(* IEC 61131-3 sources: daoli-st-library/DL_Motion, 205 files *)

(* ---- FB_DL_AxisBacklashIdent.st ---- *)
(*==============================================================================
 * 组件名称 (Component)  : FB_DL_AxisBacklashIdent
 * 所属子库 (Sublibrary) : DL_Motion
 * 当前版本 (Version)    : 1.0.0
 * 兼容性   (Platform)   : CODESYS 3.5+ / TwinCAT 3 / 汇川 InoProShop / 施耐德 Machine Expert
 *                         仅依赖 Standard.library（R_TRIG），零厂商私有库
 * 功能描述 (Function)   : 反向间隙在线辨识（只辨识、不注入）。
 *                         原理：换向瞬间传动链要"先吃掉间隙"才带动负载，故换向后的**指令位移**与
 *                         **实际位移**之差即间隙的一次观测值。本件在每个换向沿开启一个位移窗，
 *                         窗内位移超过 fWinMoveMm 即结算一个残差样本：
 *                           残差 = | (Δ指令位移) − (Δ实际位移) | [mm]
 *                         样本进定长缓冲（8 个），样本数达 nMinSamples 后取**中值**作为间隙估计
 *                         （中值对个别打滑/编码器毛刺样本免疫，均值则不）。
 *                         三条固化纪律：
 *                           ① **激励不足拒辨识**：样本数不足或换向时速度幅值低于 fVelMin 时，
 *                              估计值不宣称（bValid=FALSE）并置 bInsufficientExc——低速换向的残差
 *                              被摩擦完全淹没，硬算出来的"间隙"只是摩擦的另一种写法；
 *                           ② **中值估计**：样本排序后取中位（8 个样本插入排序，循环上界恒定）；
 *                           ③ **估计值钳位**：结果钳 [0, fBacklashMax]，超上限按上限报告并置 bClamped
 *                              （不可信的巨值不许直接进入补偿环节）。
 *                         验收向量：
 *                           ① 五次换向残差 {0.02, 0.03, 0.03, 0.04, 0.10} → 中值 0.03 mm（0.10 为野值）
 *                           ② 仅 2 个样本（nMinSamples=5）→ bValid=FALSE + bInsufficientExc
 *                           ③ 换向时速度 0.5 mm/s（fVelMin=2.0）→ 该次不采样本
 *                           ④ 残差 5.0 mm（上限 2.0）→ 估计钳 2.0 mm + bClamped
 * 接口     (Interface)  : 入 bEnable 使能、fCmdPos 指令位置、fActPos 实际位置、fVelCmd 指令速度、
 *                         fVelMin 换向速度下限（激励门槛）、fWinMoveMm 位移窗宽、fBacklashMax 估计上限、
 *                         nMinSamples 最少样本数（≥1）、bClear 清样本沿、bReset 复位沿；
 *                         出 fBacklashMm 间隙估计（中值）、bValid 估计有效、bClamped 估计被钳位、
 *                         iSampleCnt 已收样本数、bInsufficientExc 激励不足、bReversed 换向脉冲（单拍）、
 *                         eState 相、eCause 成因、bError 故障标志。
 * 边界     (Boundary)   : ① **属主边界（写死）：本件只做"间隙辨识"，不注入补偿、不改位置环输出**——
 *                         补偿注入属上层（`FB_DL_AxisCoggingFf` 族与本件并列不互引）；
 *                         ② **状态枚举禁定义**：本件不引用任何轴状态枚举（R277），只消费位置/速度引脚；
 *                         ③ **组态闸**：fVelMin > 0、fWinMoveMm > 0、fBacklashMax > 0、nMinSamples ≥ 1
 *                         且 ≤ 8，违反即锁存 eCfgIllegal；
 *                         ④ **非有限闸**：任一位置/速度样本非有限 → 该拍不采样（不锁存）；
 *                         ⑤ **样本缓冲边界**：8 样本字面量上界（R104），写入前判满；
 *                         ⑥ **锁存解除式**：eFault 仅由 bReset 上升沿解除（R228B），bReset 恒可达；
 *                         ⑦ 零全局耦合、零物理地址。
 * 分工声明 (Scope)      : 本件只管"换向残差统计与中值估计"。不接管：摩擦前馈
 *                         （属 FB_DL_AxisFrictionFf）、齿槽前馈（属 FB_DL_AxisCoggingFf）、
 *                         双反馈切换（属 AxisFeedbackFailoverSeq 族）。
 * 来源标签 (Source Tag) : 自研线（传动精度族开族）
 * 码表     (Codes)      : 本件不占用任何全局数字码位（零码位范式 R297）；诊断由 BOOL + ENUM 出口承担。
 * 红线自检 (Redline)    : R1 ✓ 零 GVL/VAR_EXTERNAL ｜ R2 ✓ 零 %I/%Q/%M ｜ R3 ✓ 纯 IEC 61131-3
 *                         R4 ✓ 组态闸 + 非有限闸 + 缓冲边界 + 估计钳位 ｜ R5 ✓ 声明逐行同行双语注释
 *                         R6 ✓ ENUM+CASE 含 ELSE 兜底 ｜ R7 ✓ 三 R_TRIG 段 0 无条件刷新（本件无 TON）
 * 修订历史 (Revision)   : 2026-11-19  v1.0.0  R47 首版（批次 4 · 序号 19）
 *==============================================================================*)

TYPE E_DL_AbiState :
(
    eIdle  := 0,    // 待机相（未使能或已清零） / Idle, disabled or cleared
    eWatch := 10,   // 观测相（等换向沿并结算样本） / Watching, awaiting reversal and sample settlement
    eFault := 90    // 故障相（组态非法，等复位） / Fault, awaiting reset
);
END_TYPE

TYPE E_DL_AbiCause :
(
    eNone           := 0,   // 无异常 / No anomaly
    eCfgIllegal     := 1,   // 组态非法（门槛/窗口/上限/样本数越域） / Illegal configuration
    eInsufficientExc:= 2,   // 激励不足（样本数不够或换向速度过低） / Insufficient excitation
    eClamped        := 3,   // 估计值被钳位（野值） / Estimate clamped
    eSampleBad      := 4,   // 位置/速度样本非有限（当拍不采） / Non-finite sample, skipped
    ePhaseBad       := 5    // 非法相位兜底 / Illegal phase fallback
);
END_TYPE

FUNCTION_BLOCK FB_DL_AxisBacklashIdent
VAR_INPUT
    bEnable      : BOOL := FALSE;      // 使能（FALSE 冻结观测，不宣称） [-] / Enable
    fCmdPos      : LREAL := 0.0;       // 指令位置 [mm] / Command position [mm]
    fActPos      : LREAL := 0.0;       // 实际位置 [mm] / Actual position [mm]
    fVelCmd      : LREAL := 0.0;       // 指令速度（用于换向判定） [mm/s] / Command velocity [mm/s]
    fVelMin      : LREAL := 2.0;       // 换向速度下限（激励门槛），域 > 0 [mm/s] / Reversal speed limit, > 0
    fWinMoveMm   : LREAL := 1.0;       // 位移窗宽，域 > 0 [mm] / Displacement window, > 0
    fBacklashMax : LREAL := 2.0;       // 估计上限，域 > 0 [mm] / Estimate ceiling, > 0
    nMinSamples  : INT := 5;           // 最少样本数，域 1..8 [个] / Minimum sample count, 1..8
    bClear       : BOOL := FALSE;      // 清样本沿（重新辨识） [-] / Clear-samples edge
    bReset       : BOOL := FALSE;      // 故障复位沿 [-] / Fault reset edge
END_VAR
VAR_OUTPUT
    fBacklashMm   : LREAL := 0.0;                        // 间隙估计（中值，已钳位） [mm] / Backlash estimate, clamped
    bValid        : BOOL := FALSE;                       // 估计有效（样本够且激励足） [-] / Estimate valid
    bClamped      : BOOL := FALSE;                       // 估计被钳位 [-] / Estimate clamped
    iSampleCnt    : INT := 0;                            // 已收样本数 [个] / Collected sample count
    bInsufficientExc : BOOL := FALSE;                    // 激励不足 [-] / Insufficient excitation
    bReversed     : BOOL := FALSE;                       // 换向脉冲（单拍） [-] / Reversal pulse, single scan
    eState        : E_DL_AbiState := E_DL_AbiState.eIdle;    // 相出口 [-] / Phase outlet
    eCause        : E_DL_AbiCause := E_DL_AbiCause.eNone;    // 成因出口（R190 归因唯一） [-] / Cause outlet
    bError        : BOOL := FALSE;                       // 故障标志（仅组态级） [-] / Error flag, configuration only
END_VAR
VAR
    _eState   : E_DL_AbiState := E_DL_AbiState.eIdle;    // 内部相（CASE 唯一写入目标） / Internal phase
    _eCause   : E_DL_AbiCause := E_DL_AbiCause.eNone;    // 成因锁存量 / Latched cause
    _bFault   : BOOL := FALSE;                           // 故障锁存位 / Latched fault bit
    _iCnt     : INT := 0;                                // 样本计数 / Sample count
    _bDirPos  : BOOL := FALSE;                           // 上拍方向为正标志 / Previous direction positive flag
    _bDirNow  : BOOL := FALSE;                           // 当拍方向标志 / Present direction flag
    _bWinOpen : BOOL := FALSE;                           // 位移窗开启标志 / Displacement window open
    _fCmdSnap : LREAL := 0.0;                            // 换向瞬间指令位置快照 [mm] / Command snapshot at reversal
    _fActSnap : LREAL := 0.0;                            // 换向瞬间实际位置快照 [mm] / Actual snapshot at reversal
    _fResid   : LREAL := 0.0;                            // 残差工作值 [mm] / Residual working value
    _fEst     : LREAL := 0.0;                            // 中值估计工作值 [mm] / Median working value
    _fTmp     : LREAL := 0.0;                            // 排序交换临时量 [mm] / Sort swap temporary
    _bRev     : BOOL := FALSE;                           // 换向脉冲内部位（单拍） / Internal reversal pulse
    _bClamped : BOOL := FALSE;                           // 钳位标志内部位 / Internal clamp flag
    _bSampleOk: BOOL := FALSE;                           // 样本有限性结论 / Sample finiteness result
    _bCfgBad  : BOOL := FALSE;                           // 组态非法当拍量 / Illegal configuration this scan
    _i        : INT := 0;                                // 样本循环下标 / Sample loop index
    _j        : INT := 0;                                // 排序内层下标 / Inner sort index
    rtClear   : R_TRIG;                                  // 清样本沿实例，段 0 无条件调用 / Clear edge instance
    rtReset   : R_TRIG;                                  // 复位沿实例，段 0 无条件调用 / Reset edge instance
    afSmp     : ARRAY[1..8] OF LREAL;                    // 残差样本缓冲（字面量上界，R104） [mm] / Residual sample buffer
    afSort    : ARRAY[1..8] OF LREAL;                    // 排序副本 [mm] / Sorting copy
END_VAR
VAR CONSTANT
    DL_ABI_NMAX : INT := 8;            // 样本缓冲深度（与数组字面量上界同源） [个] / Sample buffer depth
    DL_ABI_EPS  : LREAL := 1.0E-12;    // 浮点判等容差 [mm] / Equality tolerance
END_VAR

(* —— 段 0：组态闸 + 三沿无条件周期刷新（R228A；本件无 TON） —— *)
_bCfgBad := (fVelMin <= 0.0) OR (fWinMoveMm <= 0.0) OR (fBacklashMax <= 0.0)      // 三正域闸 / Three positive-domain gates
         OR (nMinSamples < 1) OR (nMinSamples > DL_ABI_NMAX);                     // 样本数域闸 / Sample count domain
rtClear(CLK := bClear);                                                            // 清样本沿 / Clear edge
rtReset(CLK := bReset);                                                            // 复位沿 / Reset edge

(* —— 段 1：单拍/输出量预置（锁存量 _eCause/_bFault/_iCnt/_bWinOpen/_bDirPos 不入清单，R107） —— *)
bValid   := FALSE;                                                                 // 有效位预置 / Validity preset
_bRev    := FALSE;                                                                 // 换向脉冲预清 / Reversal pulse preset
_bClamped:= FALSE;                                                                 // 钳位标志预清 / Clamp flag preset
bInsufficientExc := FALSE;                                                         // 激励不足预清 / Insufficient-excitation preset
bError   := FALSE;                                                                 // 故障标志预清（R45 配对） / Error preset
_fEst    := 0.0;                                                                   // 估计工作值预置 / Estimate preset

(* —— 段 2：组态闸（非法即锁存） —— *)
IF _bCfgBad THEN
    _eCause := E_DL_AbiCause.eCfgIllegal;                                          // 归因：组态非法 / Cause: illegal configuration
    _bFault := TRUE;                                                               // 锁存 / Latch
    _eState := E_DL_AbiState.eFault;                                               // 入故障相 / Enter fault phase
END_IF

(* —— 段 3：迁出链与清样本链（两条显式写出） —— *)
IF rtReset.Q THEN
    _bFault   := FALSE;                                                            // 清故障锁存 / Clear fault latch
    _eCause   := E_DL_AbiCause.eNone;                                              // 清成因 / Clear cause
    _iCnt     := 0;                                                                // 样本清零 / Samples cleared
    _bWinOpen := FALSE;                                                            // 关窗 / Window closed
    _eState   := E_DL_AbiState.eIdle;                                              // 回待机相 / Back to idle
END_IF
IF rtClear.Q THEN
    _iCnt     := 0;                                                                // 样本清零（重新辨识） / Samples cleared for re-identification
    _bWinOpen := FALSE;                                                            // 关窗 / Window closed
END_IF

(* —— 段 4：相迁移（使能驱动；故障相由段 3 迁出） —— *)
CASE _eState OF

E_DL_AbiState.eIdle:
    IF bEnable AND (NOT _bCfgBad) THEN
        _eState := E_DL_AbiState.eWatch;                                           // 使能进观测相 / Enter watching
    END_IF

E_DL_AbiState.eWatch:
    IF NOT bEnable THEN
        _eState := E_DL_AbiState.eIdle;                                            // 失能回待机相（不借故障相过桥，R211） / Back to idle
    END_IF

E_DL_AbiState.eFault:
    ;                                                                              // 故障相：由段 3 复位沿迁出 / Exit via the reset edge

ELSE
    _eCause := E_DL_AbiCause.ePhaseBad;                                            // 归因：非法相位 / Cause: illegal phase
    _bFault := TRUE;                                                               // 锁存 / Latch
    _eState := E_DL_AbiState.eFault;                                               // 强拉故障相 / Force fault phase

END_CASE

(* —— 段 5：换向检测与窗结算（样本采集唯一入口） —— *)
IF _eState = E_DL_AbiState.eWatch THEN
    _bSampleOk := NOT ((fCmdPos <> fCmdPos) OR ((fCmdPos - fCmdPos) <> (fCmdPos - fCmdPos)))
              AND NOT ((fActPos <> fActPos) OR ((fActPos - fActPos) <> (fActPos - fActPos)))
              AND NOT ((fVelCmd <> fVelCmd) OR ((fVelCmd - fVelCmd) <> (fVelCmd - fVelCmd)));

    IF _bSampleOk THEN
        (* 换向判定：速度符号翻转且幅值过激励门槛；方向保持量只在激励充分时更新 *)
        _bDirNow := (fVelCmd > 0.0);                                               // 本拍方向 / Present direction
        IF (ABS(fVelCmd) > fVelMin) THEN
            IF (_bDirNow <> _bDirPos) AND (NOT _bWinOpen) THEN
                _bRev     := TRUE;                                                 // 换向脉冲（内部位） / Internal reversal pulse
                _bWinOpen := TRUE;                                                 // 开位移窗 / Open the displacement window
                _fCmdSnap := fCmdPos;                                              // 记录指令基准 / Command snapshot
                _fActSnap := fActPos;                                              // 记录实际基准 / Actual snapshot
            END_IF
            _bDirPos := _bDirNow;                                                  // 方向保持量更新 / Refresh the direction
        END_IF

        (* 窗结算：指令位移超过窗宽即结算一个残差样本 *)
        IF _bWinOpen AND (ABS(fCmdPos - _fCmdSnap) > fWinMoveMm) THEN
            _fResid := ABS((fCmdPos - _fCmdSnap) - (fActPos - _fActSnap));         // 残差 = |Δ指令 − Δ实际| / Residual
            IF _fResid <> _fResid THEN
                _fResid := 0.0;                                                    // 残差非有限：拒收（不采样本） / Non-finite residual rejected
                _eCause := E_DL_AbiCause.eSampleBad;                               // 归因：样本非有限 / Cause: sample non-finite
            ELSIF _iCnt < DL_ABI_NMAX THEN
                _iCnt := _iCnt + 1;                                                // 样本计数 +1 / Sample count increment
                afSmp[_iCnt] := _fResid;                                           // 落样本（下标已判满） / Store the sample
            END_IF
            _bWinOpen := FALSE;                                                    // 关窗，等下次换向 / Close the window
        END_IF
    ELSE
        _eCause := E_DL_AbiCause.eSampleBad;                                       // 归因：样本非有限（当拍不采） / Cause: non-finite sample
    END_IF

    (* —— 段 6：中值估计（只对已收样本排序；插入排序，循环上界为样本数 ≤ 8） —— *)
    IF _iCnt >= nMinSamples THEN
        FOR _i := 1 TO _iCnt DO
            afSort[_i] := afSmp[_i];                                               // 复制已收样本 / Copy the collected samples
        END_FOR
        FOR _i := 2 TO _iCnt DO
            _j := _i;                                                              // 插入排序内层起点 / Insertion start
            WHILE (_j > 1) AND (afSort[_j - 1] > afSort[_j]) DO
                _fTmp := afSort[_j - 1];                                           // 交换 / Swap
                afSort[_j - 1] := afSort[_j];
                afSort[_j] := _fTmp;
                _j := _j - 1;                                                      // 内层推进（收敛，R74） / Inner step, converges
            END_WHILE
        END_FOR
        _fEst := afSort[(_iCnt / 2) + 1];                                          // 取中位（1 基，样本数 1..8） / Median, 1-based
        IF _fEst > fBacklashMax THEN
            _fEst := fBacklashMax;                                                 // 上限钳位（野值不许进入补偿） / Clamp to the ceiling
            _bClamped := TRUE;                                                     // 钳位标志 / Clamp flag
            _eCause := E_DL_AbiCause.eClamped;                                     // 归因：估计被钳位 / Cause: estimate clamped
        ELSIF _fEst < 0.0 THEN
            _fEst := 0.0;                                                          // 下限钳位（间隙非负） / Clamp to zero
            _bClamped := TRUE;                                                     // 钳位标志 / Clamp flag
            _eCause := E_DL_AbiCause.eClamped;                                     // 归因：估计被钳位 / Cause: estimate clamped
        END_IF
        bValid := TRUE;                                                            // 估计有效 / Estimate valid
    ELSE
        bInsufficientExc := TRUE;                                                  // 激励不足：不宣称 / Insufficient excitation
        _eCause := E_DL_AbiCause.eInsufficientExc;                                 // 归因：激励不足 / Cause: insufficient excitation
    END_IF
END_IF

(* —— 段 7：出口单点映射（名实双出口，R191） —— *)
fBacklashMm := _fEst;                                                              // 间隙估计出口 / Backlash estimate outlet
bClamped    := _bClamped;                                                          // 钳位标志出口 / Clamp flag outlet
iSampleCnt  := _iCnt;                                                              // 样本数出口 / Sample count outlet
bReversed   := _bRev;                                                              // 换向脉冲出口 / Reversal pulse outlet
eState      := _eState;                                                            // 相出口 / Phase outlet
eCause      := _eCause;                                                            // 成因出口 / Cause outlet
bError      := _bFault;                                                            // 故障标志 / Error flag

END_FUNCTION_BLOCK

(* ---- FB_DL_AxisFeedbackFailoverSeq.st ---- *)
(*==============================================================================
 * 组件名称 (Component)  : FB_DL_AxisFeedbackFailoverSeq
 * 所属子库 (Sublibrary) : DL_Motion
 * 当前版本 (Version)    : 1.0.1
 * 兼容性   (Platform)   : CODESYS 3.5+ / TwinCAT 3 / 汇川 InoProShop / 施耐德 Machine Expert
 *                         仅依赖 Standard.library（TON / R_TRIG / ABS），零厂商私有库
 * 功能描述 (Function)   : 主反馈（负载侧光栅尺/全闭环编码器）失效 → 电机侧反馈降级切换序。
 *                         四段序，每段语义显式，绝无"静默降级"：
 *                           ① ePrimary 主用相：bUsePrimary=TRUE，主反馈在岗；
 *                           ② eConfirm 失主确认相：主反馈有效位为假且持续 tLossConfirm；
 *                           ③ eSwitching 切换过渡相：**两侧均不宣称可用**（bUsePrimary 与
 *                              bUseMotorSide 同为假），先撤主用再等 tSwitchDwell，让轴级看到
 *                             一个明确的"无有效反馈"过渡拍，禁止无缝瞬切造成位置基准跳变；
 *                           ④ eDegraded 降级保持相：bUseMotorSide=TRUE 且 bFailoverActive 锁存置真，
 *                             告警持续可见直到人工复位（不因主反馈恢复而自动消失——那会让
 *                             维护人员永远看不到发生过降级）。
 *                         另设 eBlocked：主反馈已失效但 bSwitchPermit 为假（轴在运动中、
 *                         未到安全位）→ 置 bSwitchForbidden 告警，两侧反馈出口同为假，
 *                         交由轴级停机；**不做"先切了再说"**。
 * 接口     (Interface)  : 输入 bPrimaryValid 主反馈有效位、bSwitchPermit 允许切换（安全前置）、
 *                         tLossConfirm 失主确认时间、tSwitchDwell 切换过渡驻留时间、bReset 复位；
 *                         输出 bUsePrimary 用主反馈、bUseMotorSide 用电机侧、bFailoverActive
 *                         降级告警锁存、bSwitchForbidden 切换被禁止告警、eState / eCause / bError。
 * 边界     (Boundary)   : ① **属主边界（写死）：本件是"切换序"的唯一属主**——它决定何时撤主用、
 *                         何时上电机侧、过渡驻留多久。**判"负载侧是否可信"不是本件的职责**，
 *                         那属于 `FB_DL_AxisLoadEncoderLossMonitor`；本件只吃它的结论位
 *                         bPrimaryValid，不得内嵌断线/冻结判据（否则两件归因冲突、故障台账双记）。
 *                         ② 本件**不使能/不停止轴、不发运动指令**，只出反馈选择与告警位，
 *                         降级后的速度/位置环怎么跑由轴级 POU 决定。
 *                         ③ 组态闸：tLossConfirm <= T#0S → 故障锁存（防零时切换）。tSwitchDwell 的
 *                            "域 >= T#0S" 由类型本身保证（TIME 无符号），v1.0.1 已删除该恒假判据。
 *                         ④ 两枚 TON + 一枚 R_TRIG 段 0 无条件周期刷新，PT 语义成对写死；
 *                         切换过渡用 tonDwell（IN = 当拍位于 eSwitching），出相即 IN 落假自动复位，
 *                         无跨相累积（R228A）。
 *                         ⑤ 故障相与降级相均可迁出（R228B）：bReset 上升沿 → ePrimary。
 *                         ⑥ 零全局耦合（无 GVL / 无 VAR_EXTERNAL / 无物理地址）。
 * 分工声明 (Scope)      : 与 `FB_DL_AxisLoadEncoderLossMonitor`（只判负载侧可信度）、
 *                         `FB_DL_AxisDualFeedbackGuard`（双侧交叉校核）三件成组：监控件出结论，
 *                         本件按结论执行切换，校核件做一致性体检。三件互不内嵌对方判据。
 * 来源标签 (Source Tag) : P1 双反馈族 / T2-4 ◐
 * 解除式   (Release)    : bReset 上升沿（人工确认）→ 回 ePrimary 并清 bFailoverActive。
 *                         自证可满足：复位是外部操作员动作，不受任何锁存量门控；不设"主反馈自动
 *                         恢复即回切"的隐式路径——那会在反馈抖动时来回切换，且会抹掉降级告警痕迹。
 * 码表     (Codes)      : 本件不占用任何全局数字码位。出口为 BOOL（bUsePrimary / bUseMotorSide /
 *                         bFailoverActive / bSwitchForbidden / bError）+ ENUM（eState / eCause）；
 *                         数字码位待主控收口阶段统一派号（R46 码位规则）。
 * 红线自检 (Redline)    : R1 ✓ 零 GVL/VAR_EXTERNAL ｜ R2 ✓ 零 %I/%Q/%M ｜ R3 ✓ 纯 IEC 61131-3
 *                         R4 ✓ 时间域几何闸 + 无浮点比较 ｜ R5 ✓ 声明逐行同行双语注释
 *                         R6 ✓ ENUM+CASE 含 ELSE ｜ R7 ✓ TON/R_TRIG 段 0 无条件刷新
 * 返修记录 (Repair)     : v1.0.1（R47 P0 返修）① bError 出口增 `(_eState = eFault)` 项——原先只有禁止相
 *                         置位，故障相虽锁存却不报错，轴级不会停机；② 删除 `tSwitchDwell < T#0S` 恒假死检查
 *                         （TIME 为无符号时长量，与 0 的"小于"结构性不可达，属死判据）。
 * 修订历史 (Revision)   : 2026-11-19  v1.0.0  R46 首版（批次 2 · 序号 6）
 *==============================================================================*)

TYPE E_DL_FfsState :
(
    ePrimary   := 0,    // 主反馈在岗相 / Primary feedback in service
    eConfirm   := 10,   // 失主确认相（等 tLossConfirm） / Primary-loss confirmation
    eSwitching := 20,   // 切换过渡相（两侧均不宣称可用） / Switching transition, neither side claimed
    eDegraded  := 30,   // 降级保持相（电机侧在岗，告警锁存） / Degraded hold, alarm latched
    eBlocked   := 40,   // 切换被禁止相（安全前置未满足） / Switch forbidden phase
    eFault     := 90    // 组态故障相 / Configuration fault phase
);
END_TYPE

TYPE E_DL_FfsCause :
(
    eNone           := 0,   // 无故障成因 / No cause
    eCfgIllegal     := 1,   // 组态非法（确认时间非正/驻留为负） / Illegal configuration
    ePrimaryLost    := 2,   // 主反馈失效并已确认，完成降级 / Primary lost and confirmed, degraded
    eSwitchForbidden:= 3,   // 主反馈失效但切换前置不满足 / Primary lost but switching not permitted
    ePhaseBad       := 4    // 非法相位兜底 / Illegal phase fallback
);
END_TYPE

FUNCTION_BLOCK FB_DL_AxisFeedbackFailoverSeq
VAR_INPUT
    bPrimaryValid  : BOOL := TRUE;          // 主反馈（负载侧）有效位，来自监控件 [-] / Primary feedback validity, from the monitor unit
    bSwitchPermit  : BOOL := FALSE;         // 允许切换的安全前置（轴静止/在安全位） [-] / Safety precondition permitting the switch
    tLossConfirm   : TIME := T#100MS;       // 失主确认时间，域 > T#0S [ms] / Primary-loss confirm time, domain > T#0S
    tSwitchDwell   : TIME := T#20MS;        // 切换过渡驻留时间，域 >= T#0S [ms] / Switching dwell, domain >= T#0S
    bReset         : BOOL := FALSE;         // 人工复位，上升沿回主用相并清降级告警 [-] / Manual reset, rising edge returns to primary
END_VAR
VAR_OUTPUT
    bUsePrimary     : BOOL;     // 采用主反馈（负载侧） [-] / Use primary feedback
    bUseMotorSide   : BOOL;     // 采用电机侧反馈（降级后） [-] / Use motor-side feedback
    bFailoverActive : BOOL;     // 降级告警，锁存保持到复位（显式，不静默） [-] / Failover alarm, latched until reset
    bSwitchForbidden: BOOL;     // 切换被禁止告警（当拍量） [-] / Switch-forbidden alarm, per scan
    eState          : E_DL_FfsState;    // 状态出口 [-] / State outlet
    eCause          : E_DL_FfsCause;    // 成因出口（R190 归因唯一） [-] / Cause outlet
    bError          : BOOL;             // 故障标志（组态故障或切换被禁止） [-] / Error flag
END_VAR
VAR
    _eState    : E_DL_FfsState := E_DL_FfsState.ePrimary;    // 内部相位（CASE 唯一写入目标） / Internal phase
    _eCause    : E_DL_FfsCause := E_DL_FfsCause.eNone;       // 成因出口暂存（锁存语义由相位承载） / Cause staging
    tonLoss    : TON;           // 失主确认计时，段 0 无条件调用 / Primary-loss confirm timer
    tonDwell   : TON;           // 切换过渡驻留计时，段 0 无条件调用 / Switching dwell timer
    rtReset    : R_TRIG;        // 复位沿实例，段 0 无条件调用 / Reset edge instance
    _bFailover : BOOL;          // 降级告警锁存位（锁存量，仅复位沿清） / Latched failover alarm
    _bCfgBad   : BOOL;          // 组态非法当拍量 [-] / Illegal configuration this scan
END_VAR

(* —— 段 0：判据派生 + 两 TON 一沿无条件周期刷新 —— *)
_bCfgBad := (tLossConfirm <= T#0S);                             // 时间域几何闸（v1.0.1 删 tSwitchDwell < T#0S 恒假判据：TIME 无符号） / Time-domain geometry gate
rtReset(CLK := bReset);                                          // 复位沿，每拍必调（R228A） / Reset edge, every scan
tonLoss(IN := NOT bPrimaryValid, PT := tLossConfirm);            // 失主确认：有效位为假即计时（IN 由当拍判据派生） / Loss confirm, IN derived per scan
tonDwell(IN := (_eState = E_DL_FfsState.eSwitching), PT := tSwitchDwell);   // 过渡驻留：仅在过渡相计时，出相自复位 / Dwell only in transition phase

(* —— 段 1：单拍量预清零（锁存量 _bFailover / _eCause 不入清单，R107） —— *)
bUsePrimary      := FALSE;      // 主用出口每拍预清 / Primary outlet preset
bUseMotorSide    := FALSE;      // 电机侧出口每拍预清 / Motor-side outlet preset
bFailoverActive  := FALSE;      // 降级告警每拍预清，锁存分支同拍回填 / Failover alarm preset
bSwitchForbidden := FALSE;      // 禁止切换告警每拍预清 / Forbidden alarm preset
bError           := FALSE;      // 故障标志每拍预清（R45 配对） / Error flag preset

(* —— 段 2：复位沿（唯一回主用路径，人工确认语义） —— *)
IF rtReset.Q THEN
    _bFailover := FALSE;                    // 清降级告警锁存（锁存量） / Clear latched failover alarm
    _eCause    := E_DL_FfsCause.eNone;      // 清成因 / Clear cause
    _eState    := E_DL_FfsState.ePrimary;   // 回主用相（R228B 迁出路径） / Return to primary phase
END_IF

(* —— 段 3：组态闸（先于相位机，保证每拍一致） —— *)
IF _bCfgBad THEN
    _eState := E_DL_FfsState.eFault;        // 组态非法入故障相 / Enter fault phase
    _eCause := E_DL_FfsCause.eCfgIllegal;   // 归因：组态非法 / Cause: illegal configuration
    bError  := TRUE;                        // 故障标志同拍置位 / Error flag set same scan
END_IF

(* —— 段 4：相位机（ENUM 全成员显式标签 + ELSE 兜底，R128） —— *)
CASE _eState OF

E_DL_FfsState.ePrimary:
    IF bPrimaryValid = FALSE THEN                       // 出口 1：主反馈报失效 → 进确认相（不立即切） / Primary reported invalid, confirm first
        _eState := E_DL_FfsState.eConfirm;
    ELSIF rtReset.Q THEN                                // 出口 2：复位沿保持主用相（幂等） / Reset keeps primary, idempotent
        _eState := E_DL_FfsState.ePrimary;
    END_IF

E_DL_FfsState.eConfirm:
    IF bPrimaryValid THEN                               // 出口 1：有效位回真（抖动）→ 回主用，不留痕 / Validity returned, back to primary without a trace
        _eState := E_DL_FfsState.ePrimary;
    ELSIF tonLoss.Q THEN                                // 出口 2：确认窗到 → 看安全前置 / Confirm window elapsed, check precondition
        IF bSwitchPermit THEN
            _eState := E_DL_FfsState.eSwitching;        // 前置满足：进切换过渡 / Precondition met, enter transition
        ELSE
            _eState := E_DL_FfsState.eBlocked;          // 前置不满足：进禁止相（不硬切） / Precondition unmet, forbid the switch
        END_IF
    END_IF

E_DL_FfsState.eSwitching:
    IF rtReset.Q THEN                                   // 出口 1：过渡中人工复位 → 回主用相 / Reset during transition
        _eState := E_DL_FfsState.ePrimary;
    ELSIF NOT bSwitchPermit THEN                        // 出口 2：前置撤销（轴动起来了）→ 撤回并进禁止相 / Precondition withdrawn
        _eState := E_DL_FfsState.eBlocked;
    ELSIF tonDwell.Q THEN                               // 出口 3：驻留到 → 上电机侧并锁存告警 / Dwell elapsed, engage motor side
        _bFailover := TRUE;                             // 告警锁存（锁存量） / Latch the alarm
        _eCause    := E_DL_FfsCause.ePrimaryLost;       // 归因：主反馈失效已完成降级 / Cause: primary lost, degraded
        _eState    := E_DL_FfsState.eDegraded;
    END_IF

E_DL_FfsState.eDegraded:
    IF rtReset.Q THEN                                   // 出口：仅人工复位可离开降级相 / Only a manual reset leaves degradation
        _eState := E_DL_FfsState.ePrimary;
    END_IF

E_DL_FfsState.eBlocked:
    IF bPrimaryValid THEN                               // 出口 1：主反馈自己回来了 → 回主用（解除禁止） / Primary recovered by itself
        _eState := E_DL_FfsState.ePrimary;
    ELSIF bSwitchPermit AND tonLoss.Q THEN              // 出口 2：前置满足且确认仍在 → 进切换过渡 / Precondition now met
        _eState := E_DL_FfsState.eSwitching;
    END_IF

E_DL_FfsState.eFault:
    IF rtReset.Q AND (NOT _bCfgBad) THEN                // 出口：复位沿 + 组态已合法才迁出（R228B） / Reset edge with legal config
        _eState := E_DL_FfsState.ePrimary;
    END_IF

ELSE
    _eCause := E_DL_FfsCause.ePhaseBad;                 // 归因：非法相位 / Cause: illegal phase
    _eState := E_DL_FfsState.eFault;                    // 强拉故障相 / Force fault phase
    bError  := TRUE;                                    // 故障标志 / Error flag

END_CASE

(* —— 段 5：出口单点映射（名实同源；过渡相两侧皆假是设计意图，非缺省） —— *)
CASE _eState OF
E_DL_FfsState.ePrimary:
    bUsePrimary := TRUE;                                // 主用相：取主反馈 / Primary phase uses primary feedback
E_DL_FfsState.eDegraded:
    bUseMotorSide := TRUE;                              // 降级相：取电机侧 / Degraded phase uses motor side
E_DL_FfsState.eBlocked:
    bSwitchForbidden := TRUE;                           // 禁止相：显式告警 / Forbidden phase raises the alarm
    bError           := TRUE;                           // 禁止相属故障级（轴级据此停机） / Forbidden is fault level
ELSE
    ;                                                   // 其余相（确认/过渡/故障）：两侧均不宣称可用 / Other phases claim neither side
END_CASE
bFailoverActive := _bFailover;                          // 降级告警与锁存同源（R191） / Alarm from latch
bError          := bError OR (_eState = E_DL_FfsState.eFault);   // v1.0.1：故障相必置故障标志（原先仅禁止相置位） / Fault phase forces the error flag
eState          := _eState;                             // 状态出口 / State outlet
eCause          := _eCause;                             // 成因出口 / Cause outlet

END_FUNCTION_BLOCK

(* ---- FB_DL_AxisInPosMonitor.st ---- *)
(*
    FB_DL_AxisInPosMonitor —— 到位稳定判定
    ------------------------------------------------------------------
    分类      : DL_Motion / AxisMonitor
    前缀      : FB_DL_
    版本      : 1.0.0
    溯源      : T1-6 PLCopen（只借 InPosition / Standstill 两个公开输出的语义边界：
                InPosition = 位置入窗，Standstill = 速度低于阈；两者都是「判定」而非「指令」）；
                稳定时间、抖振窗、掩码与码位 100% 自有；clean-room 重写，
                未复制任何闭源厂商源码，参考实现仅限 MIT/Apache 许可
    道莅 clean-room 防御性实现：语义借鉴、代码与码位 100% 自有
    平台      : 纯 IEC 61131-3，CODESYS V3.5+ / TwinCAT 3 / InoProShop / Machine Expert 通用
    作者      : 道莅代码库 · PLC编程专家（R22 批 4 · #16）
    ------------------------------------------------------------------
    功能说明  : 机械手取放、压装、点胶这类「必须真停稳才能动作」的工位，需要一个比驱动器
                内置信号更严的到位判据：位置进窗 + 速度进阈 + 连续稳定满 tSettle 才算到位。
                本件就地给出三层结论——瞬时入窗（bInPos）、稳定到位（bSettled，取放联锁用
                这一个）、抖振超限（bChatterAlarm，稳定窗内反复出窗说明伺服在追或机械在弹）。
    职责划界  : 驱动器内置的跟随误差监视（FB_DL_AxisFollowingErrorMonitor）看的是
                「指令位置与实际位置的偏差」是否超限，管的是伺服跟随品质与保护停机；
                本件看的是「实际位置是否已稳定落在目标窗内」，管的是工艺许可。
                两者判据不同、出口不同、处置不同：前者越限要停轴，后者越限只是不许动作。
                本件不重复实现跟随误差保护，也不发任何运动指令、不改写轴状态。
    轴故障口径: 与批 4 其余各件一致——本件不消费 bAxisError 引脚，也绝不代替轴侧做恢复动作。
                轴一旦报故障停车，判定必然出窗并自然退回 eMoving，bSettled 当拍清零；
                恢复只能由轴侧完成后重新走「入窗 → 稳定满 tSettle」，本件不做任何自动续判。
    非有限值  : 采样出现 NaN / ±Inf 时判定冻结（保持上次判定）并报 02F7，绝不拿坏值
                伪造「到位」。因此下游取放联锁必须写成「bSettled AND bValid」——
                bSettled 只是判定值，bValid 才是「这个判定值可信」的凭据（语义分离，
                二者不可互相替代）。
    边界安全  : ① 容差与时间参数非法 → 02F6、bValid = FALSE、全输出清零并进 eFault；
                ② 采样非有限 → 02F7、判定与两只定时器全部冻结，坏值消失后重新起算；
                ③ bSettled 出窗当拍即清零，绝不锁存到下一件料（R34 家族）；
                ④ 失能 → 逐项清零输出（R72 双路径：先全清再按状态置位）；
                ⑤ 抖振计数按观察窗清，窗口自重启（TON 自复位构成滚动窗）。
    错误码    : 16#0004_01DD 已入窗但稳定时间未到，暂不计到位——信息级，入稳相那一拍发布
                16#0004_01DE 抖振计数已按观察窗清零，稳定保持——信息级
                16#0004_02F6 容差或时间参数非法（容差非正 / 稳定时间为零 / 窗长为零）——故障级
                16#0004_02F7 位置或速度采样非有限，判定冻结并保持上次判定——故障级，非锁存
                16#0004_02F8 状态机落 ELSE 兜底（非法状态）——故障级
    码位总账  : 16#0004_01DD 用 / 16#0004_01DE 用 ｜ 16#0004_02F6 用 / 16#0004_02F7 用 / 16#0004_02F8 用
    状态机    : E_DL_InPosState（eIdle / eMoving / eSettling / eInPos / eChatter / eFault），
                CASE 含 ELSE 兜底，ELSE 置 16#0004_02F8 并回 eFault；失能无条件回 eIdle。
    采样约定  : fbSettle 与 fbChatterWin 在本体最前部无条件调用（R40）；窗定时器以
                「IN := NOT 自身 Q」自重启构成滚动窗，Q 只亮一拍即完成清零动作；
                段转出统一走「断输入一拍」标志，标志在对应调用之后立刻自清。
    依赖      : 仅 Standard.library（TON / ABS / MIN / MAX），不引用任何其他 DL_ 子库。
    验收向量  :
                V1 域外早退：fPosTol = 0 → 02F6、bError = TRUE、bValid = FALSE、
                   bInPos / bSettled / bChatterAlarm 全 FALSE、进 eFault。
                V2 上限/超限：位置在窗内但速度 5 mm/s > fVelTol 1.0 → bInPos = FALSE，
                   不得进入 eSettling，稳定计时不启动。
                V3 跨段时序：入窗后第 tSettle−1 拍报 01DD 且 bSettled = FALSE；
                   第 tSettle 拍 bSettled 当拍置 TRUE（不延后一拍）。
                V4 恢复/抖振：窗内反复出窗 5 次（uChatterLimit = 5）→ bChatterAlarm = TRUE、
                   进 eChatter；随后重新稳定满 tSettle → 回 eInPos 且计数清零、01DE。
                V5 坏值冻结：fActPos = NaN 一拍 → 02F7、bValid = FALSE、
                   bSettled 保持坏值前一拍的判定值不变；下一拍正常采样恢复判定。
    红线自检  : 1 全局变量声明零使用 / 外部变量访问零使用 / 物理地址零使用 —— 通过，全部量经引脚注入
                2 纯 IEC 61131-3 跨平台 —— 通过，仅 Standard.library
                3 防御性编程 —— 通过，浮点比较全部为绝对值阈或容差、无非有限穿透、无除法
                4 声明行同行中英双语注释 + 单位 —— 通过，逐行附注（含枚举成员）
                5 ENUM + CASE 且含 ELSE 兜底 —— 通过
                6 TON / R_TRIG 无条件刷新 —— 通过，段 1 两只 TON 先行调用
                7 无魔法数 —— 通过，容差与时间全部为引脚或 VAR CONSTANT
    修订记录  : 2026-11-16 v1.0.0 首次入库（R22 批 4 · #16）
*)
TYPE E_DL_InPosState :
(
    eIdle    := 0,       // 未使能或参数未就绪，全输出清零 / not enabled or parameters not ready, every output is cleared
    eMoving  := 10,      // 尚未入窗，等位置与速度同时进阈 / not yet in the window, waiting for both position and velocity
    eSettling:= 20,      // 已入窗，稳定计时中，尚不可用于取放 / inside the window and timing the settle, not yet usable by a pick-and-place
    eInPos   := 30,      // 稳定到位，bSettled 可用 / settled, bSettled may be consumed
    eChatter := 40,      // 抖振超限，观察窗内出窗次数过多 / chatter limit exceeded, too many window exits inside the observation window
    eFault   := 50       // 故障，参数非法或非法状态兜底 / fault from illegal parameters or from the fallback branch
);
END_TYPE

FUNCTION_BLOCK FB_DL_AxisInPosMonitor
VAR_INPUT
    bEnable        : BOOL;                     // 使能，FALSE 时全输出清零并回 eIdle / enable, FALSE clears every output and returns to idle
    fActPos        : REAL;                     // 轴实际位置 [mm] / axis actual position [mm]
    fTargetPos     : REAL;                     // 目标位置 [mm] / target position [mm]
    fActVel        : REAL;                     // 轴实际速度 [mm/s]，取绝对值比较 / axis actual velocity [mm/s], compared on its absolute value
    fPosTol        : REAL := 0.05;             // 位置窗半宽 [mm]，必须大于 0 / position window half-width [mm], must exceed zero
    fVelTol        : REAL := 1.0;              // 速度阈 [mm/s]，必须大于 0 / velocity threshold [mm/s], must exceed zero
    tSettle        : TIME := T#100MS;          // 稳定时间 [ms]，必须大于 0 / settle time [ms], must exceed zero
    uChatterLimit  : UINT := 5;                // 抖振计数上限 [次]，0 = 首次出窗即报警 / chatter limit [pcs], 0 alarms on the first exit
    tChatterWin    : TIME := T#2S;             // 抖振观察窗长 [ms]，必须大于 0 / chatter observation window [ms], must exceed zero
END_VAR
VAR_OUTPUT
    bInPos         : BOOL;                     // 瞬时入窗（位置在窗内且速度达标）/ instantaneously inside the window, position in band and velocity below the threshold
    bSettled       : BOOL;                     // 稳定到位，取放联锁用这个；须与 bValid 相与 / settled, used by the pick-and-place interlock, must be ANDed with bValid
    uChatterCount  : UINT;                     // 本观察窗内出窗次数 [次] / window exits inside the current observation window [pcs]
    bChatterAlarm  : BOOL;                     // 抖振报警，计数达上限置位，重新稳定后清 / chatter alarm, set when the count reaches the limit and cleared after a new settle
    eErr           : UDINT;                    // 错误码，0 表示无错 / error code, 0 means no error
    bError         : BOOL;                     // 故障级标志，仅故障级错误置位 / fault-class flag, set only on fault-level codes
    bValid         : BOOL;                     // 判定可信标志，坏值拍为 FALSE / verdict trustworthy flag, FALSE on a bad-sample scan
END_VAR
VAR
    fbSettle       : TON;                      // 稳定计时器，仅 eSettling 使用 / settle timer, used in eSettling only
    fbChatterWin   : TON;                      // 抖振观察窗定时器，自重启构成滚动窗 / chatter observation window, self-restarting to form a rolling window
    _bSettleBreak  : BOOL;                     // 稳定计时器断输入一拍标志 / break-input flag for the settle timer
    _bWinPrev      : BOOL;                     // 上一拍观察窗到期标志，用于生成窗沿 / previous-scan window expiry flag used to build the window edge
    _bInWin        : BOOL;                     // 本拍入窗条件（位置与速度同拍相与）/ in-window condition of this scan, position and velocity taken together
    _bInWinPrev    : BOOL;                     // 上一拍入窗条件，用于捕捉出窗沿 / previous-scan in-window condition used to catch the leaving edge
    _bFrozen       : BOOL;                     // 判定冻结标志，坏值拍置位 / verdict freeze flag, set on a bad-sample scan
    _uChat         : UINT;                     // 抖振计数累加器，饱和不回绕 [次] / chatter accumulator, saturating and never wrapping [pcs]
    _eState        : E_DL_InPosState;          // 当前状态 / current state
END_VAR
VAR CONSTANT
    DL_IP_UINT_MAX   : UINT := 16#FFFF;        // 抖振计数饱和上限 [次] / chatter count saturation bound [pcs]
    DL_IP_INF_GUARD  : REAL := 4.0E38;         // 非有限幅值判定阈（大于 REAL 最大值）[mm] / non-finite magnitude guard [mm]
    DL_IP_ZERO       : REAL := 0.0;            // 零值常量，避免裸字面量 [无量纲] / zero constant, avoids a bare literal [dimensionless]
    DL_IP_T_ZERO     : TIME := T#0S;           // 零时间常量，用于参数门禁 / zero time constant used by the parameter gate
END_VAR

// 段 1｜两只 TON 无条件周期刷新（红线 6：严禁放入 IF / CASE；窗定时器自重启构成滚动窗）
// segment 1, both TON instances refreshed unconditionally, the window timer restarts itself to form a rolling window
// 稳定计时器在 eSettling 与 eChatter 两相承担的是同一个物理量「连续入窗时长」，
// 不属于跨段复用；每次进相统一断输入一拍，杜绝上一相的 ET 残留。
// the settle timer measures one single quantity, the continuous in-window time, in both eSettling and eChatter,
// which is not a cross-phase reuse; every entry restarts it with one scan of a FALSE input so no elapsed time leaks.
fbSettle(IN := (((_eState = E_DL_InPosState.eSettling) OR (_eState = E_DL_InPosState.eChatter)))
             AND (NOT _bSettleBreak) AND _bInWin AND (NOT _bFrozen), PT := tSettle);
_bSettleBreak := FALSE;                         // 断输入标志用后即刻自清 / the break flag clears right after the call
fbChatterWin(IN := (NOT fbChatterWin.Q) AND bEnable, PT := tChatterWin);
// 窗到期沿：Q 只亮一拍，用上一拍 Q 构造边沿，避免边沿在本拍被清零后丢失
// the window expiry edge, Q lives for a single scan so the previous-scan Q builds the edge

// 段 2｜输出与错误状态预置 / segment 2, preset outputs and error status
eErr := 0;                                      // 预置无错误 / preset no error
bError := FALSE;                                // 预置无故障标志 / preset no error flag
bValid := TRUE;                                 // 预置判定可信 / preset the verdict as trustworthy
_bFrozen := FALSE;                              // 预置不冻结 / preset not frozen

// 段 3｜参数门禁：四条参数任一非法即不许判定（判据本身不可信，给结论就是害人）
// segment 3, the parameter gate, no verdict may be produced from untrustworthy criteria
IF (fPosTol <= DL_IP_ZERO)
   OR (fVelTol <= DL_IP_ZERO)
   OR (tSettle <= DL_IP_T_ZERO)
   OR (tChatterWin <= DL_IP_T_ZERO) THEN
    eErr := 16#0004_02F6;                       // 故障级：容差或时间参数非法 / fault: a tolerance or duration parameter is illegal
    bError := TRUE;                             // 置故障标志 / raise the fault flag
    bValid := FALSE;                            // 判定不可信 / the verdict is not trustworthy
    _bSettleBreak := TRUE;                      // 稳定计时断输入重启 / restart the settle timer
    _eState := E_DL_InPosState.eFault;          // 转故障，等参数修复后失能复位 / go to fault and wait for repaired parameters plus a disable
END_IF

// 段 4｜采样非有限检测：NaN 用自不自等捕获（该式对 ±Inf 同样成立），坏值拍整段冻结
// segment 4, non-finite detection, the self-inequality test catches NaN and infinity alike and freezes the whole scan
IF (fActPos - fActPos) <> (fActPos - fActPos) THEN
    _bFrozen := TRUE;                           // 位置采样非有限 / the position sample is not finite
ELSIF ABS(fActPos) > DL_IP_INF_GUARD THEN
    _bFrozen := TRUE;                           // 位置采样超幅值门 / the position sample exceeds the magnitude guard
ELSIF (fActVel - fActVel) <> (fActVel - fActVel) THEN
    _bFrozen := TRUE;                           // 速度采样非有限 / the velocity sample is not finite
ELSIF ABS(fActVel) > DL_IP_INF_GUARD THEN
    _bFrozen := TRUE;                           // 速度采样超幅值门 / the velocity sample exceeds the magnitude guard
ELSIF (fTargetPos - fTargetPos) <> (fTargetPos - fTargetPos) THEN
    _bFrozen := TRUE;                           // 目标位置非有限 / the target position is not finite
END_IF

IF _bFrozen THEN
    eErr := 16#0004_02F7;                       // 故障级：采样非有限，判定冻结 / fault: a non-finite sample froze the verdict
    bError := TRUE;                             // 置故障标志（非锁存，坏值消失即复位）/ raise the flag, it is not latched and drops with the bad sample
    bValid := FALSE;                            // 判定不可信，下游必须与 bSettled 相与 / the verdict is not trustworthy and must be ANDed downstream
    _bSettleBreak := TRUE;                      // 稳定计时断输入重启，绝不在坏值上计时 / restart the settle timer, nothing may mature on bad data
END_IF

// 段 5｜入窗条件与抖振计数：位置与速度同拍相与，不做先后（同拍即结论）
// segment 5, the in-window condition combines position and velocity in the same scan, and the chatter counter follows the leaving edge
_bInWin := (ABS(fActPos - fTargetPos) <= fPosTol) AND (ABS(fActVel) <= fVelTol);

IF (NOT _bFrozen) AND bEnable AND (_eState <> E_DL_InPosState.eFault) THEN
    IF _bInWinPrev AND (NOT _bInWin) THEN
        IF _uChat < DL_IP_UINT_MAX THEN
            _uChat := _uChat + 1;               // 出窗一次，计数饱和自增 / one window exit, a saturating increment
        END_IF
    END_IF
END_IF

IF fbChatterWin.Q AND (NOT _bWinPrev) THEN
    // 观察窗到期一拍：按窗清零计数；若此刻仍稳定到位，说明这一窗没有异常
    // the observation window expired, clear the count, and a still-settled state means the window was clean
    IF (_eState = E_DL_InPosState.eInPos) THEN
        eErr := 16#0004_01DE;                   // 信息级：抖振计数已按窗清零，稳定保持 / info: the count was cleared with the window and the settle holds
    END_IF
    _uChat := 0;                                // 计数按窗清零 / clear the counter with the window
END_IF
_bWinPrev := fbChatterWin.Q;                    // 更新窗到期快照 / update the window expiry snapshot
_bInWinPrev := _bInWin;                         // 更新入窗快照（坏值拍也更新，恢复后不误算一次出窗）/ update the in-window snapshot, a frozen scan updates it too so recovery does not count a phantom exit

// 段 6｜状态机：只做分类与转相，判据计算已在段 5 完成
// segment 6, the state machine classifies and switches, the criteria were computed in segment 5
IF NOT _bFrozen THEN
    CASE _eState OF
    E_DL_InPosState.eIdle:
        _uChat := 0;                            // 待机计数清零 / clear the counter while idle
        IF bEnable THEN
            _eState := E_DL_InPosState.eMoving; // 使能即开始监视 / monitoring starts with the enable
        END_IF

    E_DL_InPosState.eMoving:
        IF NOT bEnable THEN
            _uChat := 0;                        // 失能计数清零 / clear the counter when disabled
            _eState := E_DL_InPosState.eIdle;   // 回待机 / back to idle
        ELSIF _bInWin THEN
            _bSettleBreak := TRUE;              // 入窗首拍，稳定计时断输入重启 / the settle timer restarts on the entering scan
            _eState := E_DL_InPosState.eSettling;   // 进稳相 / enter the settling phase
            eErr := 16#0004_01DD;               // 信息级：已入窗但稳定时间未到 / info: inside the window but the settle time has not elapsed
        END_IF

    E_DL_InPosState.eSettling:
        IF NOT bEnable THEN
            _uChat := 0;                        // 失能计数清零 / clear the counter when disabled
            _eState := E_DL_InPosState.eIdle;   // 回待机 / back to idle
        ELSIF NOT _bInWin THEN
            _eState := E_DL_InPosState.eMoving; // 出窗，回移动相重新等 / left the window, back to moving
        ELSIF fbSettle.Q THEN
            _eState := E_DL_InPosState.eInPos;  // 稳定时间满，到位可用 / the settle time elapsed and the verdict becomes usable
        END_IF

    E_DL_InPosState.eInPos:
        IF NOT bEnable THEN
            _uChat := 0;                        // 失能计数清零 / clear the counter when disabled
            _eState := E_DL_InPosState.eIdle;   // 回待机 / back to idle
        ELSIF NOT _bInWin THEN
            _bSettleBreak := TRUE;              // 出窗即作废稳定计时，不锁存到下一条料 / the settle timing dies with the exit, never latched across a part
            IF _uChat >= uChatterLimit THEN
                _eState := E_DL_InPosState.eChatter;    // 出窗次数达上限，进抖振相 / the exits reached the limit, enter the chatter phase
            ELSE
                _eState := E_DL_InPosState.eMoving;     // 偶发出窗，回移动相 / an incidental exit, back to moving
            END_IF
        END_IF

    E_DL_InPosState.eChatter:
        IF NOT bEnable THEN
            _uChat := 0;                        // 失能计数清零 / clear the counter when disabled
            _eState := E_DL_InPosState.eIdle;   // 回待机 / back to idle
        ELSIF fbSettle.Q THEN
            _uChat := 0;                        // 重新稳定满 tSettle，抖振报警解除并清零 / a fresh settle clears both the alarm and the counter
            _eState := E_DL_InPosState.eInPos;  // 回到位相 / back to the settled phase
        END_IF

    E_DL_InPosState.eFault:
        // 退出条件：参数已修复且请求已撤——参数不修就复位只会再进故障
        // exit needs repaired parameters and a withdrawn request, a reset with bad parameters would only re-enter the fault
        IF (fPosTol > DL_IP_ZERO) AND (fVelTol > DL_IP_ZERO)
           AND (tSettle > DL_IP_T_ZERO) AND (tChatterWin > DL_IP_T_ZERO)
           AND (NOT bEnable) THEN
            _uChat := 0;                        // 计数清零 / clear the counter
            _eState := E_DL_InPosState.eIdle;   // 回待机 / back to idle
        END_IF

    ELSE
        // 非法状态兜底：绝不静默停在未知态 / illegal state fallback, never stay silently in an unknown state
        eErr := 16#0004_02F8;                   // 故障级：状态机落 ELSE / fault: the state machine fell into ELSE
        bError := TRUE;                         // 置故障标志 / raise the fault flag
        bValid := FALSE;                        // 判定不可信 / the verdict is not trustworthy
        _bSettleBreak := TRUE;                  // 稳定计时断输入重启 / restart the settle timer
        _eState := E_DL_InPosState.eFault;      // 回故障态 / go to fault
    END_CASE
END_IF

// 段 7｜输出发布（R72 双路径：逐项显式赋值，坏值拍整块不写以保持上次判定）
// segment 7, publish outputs item by item, a frozen scan writes nothing so the previous verdict survives
IF NOT _bFrozen THEN
    bInPos := _bInWin;                          // 瞬时入窗发布 / publish the instantaneous in-window condition
    bSettled := (_eState = E_DL_InPosState.eInPos);     // 稳定到位只由状态决定，出窗当拍即清零 / the settle verdict follows the state and dies on the exit scan
    bChatterAlarm := (_eState = E_DL_InPosState.eChatter);  // 抖振报警只由状态决定 / the chatter alarm follows the state
END_IF
uChatterCount := _uChat;                        // 计数发布（坏值拍也发布，计数本身未动）/ publish the counter, which is untouched on a frozen scan
END_FUNCTION_BLOCK

(* ---- FB_DL_CamDynTrim.st ---- *)
(*==============================================================================
 * 组件名称 (Component)  : FB_DL_CamDynTrim
 * 所属子库 (Sublibrary) : DL_Motion
 * 当前版本 (Version)    : 1.0.0
 * 兼容性   (Platform)   : CODESYS 3.5+ / TwinCAT 3 / 汇川 InoProShop / 施耐德 Machine Expert
 *                         仅依赖 Standard.library（ABS），零厂商私有库
 * 功能描述 (Function)   : 凸轮动态修调（相位 + 倍率双通道）：bApply 上升沿锁存
 *                         修调目标（先钳位：|fPhaseTrim| <= fPhTrimMaxDeg、
 *                         |fScaleTrim| <= fScTrimMaxPct，超幅钳位并置信息码
 *                         eClamped），生效期按 fPhRampDs/fScRampPs 斜率渐变
 *                         逼近目标（防凸轮表跳变，规格指定），双通道均到达后
 *                         bTrimActive 撤销（修调保持）；执行中（bTrimActive=
 *                         TRUE）新 bApply 沿被拒并置信息码 eBusyRej（拒绝
 *                         叠加，规格指定），拒次计数 uRejCnt。
 * 接口     (Interface)  : 输入 fPhaseTrim 相位修调请求 [deg]、fScaleTrim 倍率
 *                         修调请求 [%]、bApply 应用沿、fPhTrimMaxDeg 单次相位
 *                         修调幅值上限（域 > 0）、fScTrimMaxPct 单次倍率修调
 *                         幅值上限（域 > 0）、fPhRampDs 相位斜率（域 > 0）
 *                         [deg/s]、fScRampPs 倍率斜率（域 > 0） [%/s]、fCycle
 *                         扫描周期（<=0 用缺省） [s]、bReset 复位；输出
 *                         fPhTrimAct 生效相位修调 [deg]、fScTrimAct 生效倍率
 *                         修调 [%]、bTrimActive 斜坡执行中、uRejCnt 执行中
 *                         拒绝计数、eErrCode 错误码、bError 故障标志。
 * 边界     (Boundary)   : ① **属主边界（写死）：本件只出修调量标量对，不改写
 *                         凸轮表本体、不接管凸轮轴使能**；凸轮表插值归
 *                         `FB_DL_ElectronicCam`。
 *                         ② 生效通道单源：目标 _fPhTar/_fScTar 只在应用沿
 *                         锁存写入；生效量 _fPhAct/_fScAct 限步逼近，斜坡中
 *                         不受新请求污染（执行中拒绝叠加）。
 *                         ③ 幅值钳位：请求超上限钳到 ±上限并置信息码
 *                         eClamped（量值方向可饱和，钳位行在锁存行后置码，
 *                         先钳后码顺序无信息级丢失）。
 *                         ④ 到达判据用容差（禁浮点 =）；双通道各自独立到达，
 *                         bTrimActive = 任一通道未达。
 *                         ⑤ 组态闸：fPhTrimMaxDeg/fScTrimMaxPct/fPhRampDs/
 *                         fScRampPs 任一 <= 0 或非有限 → 锁存故障 eCfgBad，
 *                         生效量冻结保持，bTrimActive=FALSE，解除沿 = bReset
 *                         上升沿（R45 配对）。
 *                         ⑥ 零全局耦合（无 GVL / VAR_EXTERNAL / 物理地址）。
 * 分工声明 (Scope)      : 与 `FB_DL_CamPhaseTrim`/`FB_DL_CamOverrideTrim` 分工：
 *                         静态相位/倍率修调归那两件，本件为「斜坡渐生效 + 执行中
 *                         拒叠加」动态编排件；与 `FB_DL_EdgeTrimTraverse` 分工：
 *                         边缘修调归那件。
 * 来源标签 (Source Tag) : 自研线（凸轮动态修调编排为道莅防御性实现）
 * 码表     (Codes)      : 本件不占用任何全局数字码位。出口为 LREAL 修调对 +
 *                         BOOL 组 + UDINT 计数 + ENUM 错误码；数字码位待主控
 *                         收口阶段统一派号。
 * 红线自检 (Redline)    : R1 ✓ 零 GVL/VAR_EXTERNAL ｜ R2 ✓ 零 %I/%Q/%M ｜ R3 ✓ 纯 IEC 61131-3
 *                         R4 ✓ 幅值钳位 + 容差到达 + 组态锁存 + 非有限入闸
 *                         ｜ R5 ✓ 声明逐行同行双语注释
 *                         R6 N/A（锁存态无 CASE 状态机） ｜ R7 ✓ 两 R_TRIG 段 0 无条件刷新
 * 修订历史 (Revision)   : 2026-11-20  v1.0.0  R50 首版（批次 4 · 序号 19）
 * 验收向量 (Acceptance) : ① fPhTrimMaxDeg=10：请求 fPhaseTrim=15 → 钳 10，
 *                         eClamped；fPhRampDs=50, fCycle=0.01 → 单步 0.5，
 *                         20 拍达 10.0 → bTrimActive=FALSE（修调保持）；
 *                         ② 斜坡第 5 拍再发 bApply → 被拒，uRejCnt+1，
 *                         eErrCode=eBusyRej，生效量不受污染；③ fScTrimMaxPct
 *                         =0 → 锁存 eCfgBad，生效量冻结；④ bApply 请求
 *                         fPhaseTrim=3（< 上限）→ 无钳位，eOk。
 *==============================================================================*)

(*-----------------------------------------------------------------------------
 * 枚举: E_DL_CdtErr（错误码；信息级不置 bError，故障级恒伴 bError=TRUE）
 *----------------------------------------------------------------------------*)
TYPE E_DL_CdtErr :
(
    eOk      := 0,   // 正常 / Normal
    eCfgBad  := 1,   // 故障级：组态非法（上限/斜率域或非有限） / Fault: illegal configuration
    eClamped := 2,   // 信息级：请求超单次幅值上限已钳位 / Info: request clamped to single-shot ceiling
    eBusyRej := 3    // 信息级：执行中应用沿被拒（拒绝叠加） / Info: apply edge rejected while busy
);
END_TYPE

FUNCTION_BLOCK FB_DL_CamDynTrim
VAR_INPUT
    fPhaseTrim  : LREAL := 0.0;       // 相位修调请求 [deg] / Phase trim request [deg]
    fScaleTrim  : LREAL := 0.0;       // 倍率修调请求 [%] / Scale trim request [percent]
    bApply      : BOOL := FALSE;      // 应用沿（上升沿锁存目标，执行中拒绝） [-] / Apply edge
    fPhTrimMaxDeg: LREAL := 10.0;     // 单次相位修调幅值上限，域 > 0 [deg] / Single-shot phase trim ceiling
    fScTrimMaxPct: LREAL := 20.0;     // 单次倍率修调幅值上限，域 > 0 [%] / Single-shot scale trim ceiling
    fPhRampDs   : LREAL := 50.0;      // 相位斜率，域 > 0 [deg/s] / Phase ramp rate
    fScRampPs   : LREAL := 10.0;      // 倍率斜率，域 > 0 [%/s] / Scale ramp rate
    fCycle      : LREAL := 0.0;       // 扫描周期（<=0 用缺省） [s] / Scan cycle, default used when <= 0
    bReset      : BOOL := FALSE;      // 复位，上升沿清组态锁存与拒次计数 [-] / Reset, clears latch and reject counter
END_VAR
VAR_OUTPUT
    fPhTrimAct : LREAL;               // 生效相位修调（斜坡后） [deg] / Active phase trim [deg]
    fScTrimAct : LREAL;               // 生效倍率修调（斜坡后） [%] / Active scale trim [percent]
    bTrimActive: BOOL;                // 斜坡执行中指示（任一通道未达） [-] / Ramp busy indicator
    uRejCnt    : UDINT := 0;          // 执行中拒绝计数（防回绕） [次] / Busy-reject counter
    eErrCode   : E_DL_CdtErr;         // 错误码出口 / Error code outlet
    bError     : BOOL;                // 故障标志（组态锁存） [-] / Error flag, latched
END_VAR
VAR
    _fPhTar   : LREAL := 0.0;         // 相位目标锁存（应用沿唯一写入） [deg] / Phase target latch
    _fScTar   : LREAL := 0.0;         // 倍率目标锁存 [percent] / Scale target latch
    _fPhAct   : LREAL := 0.0;         // 生效相位（限步源） [deg] / Active phase internal
    _fScAct   : LREAL := 0.0;         // 生效倍率（限步源） [percent] / Active scale internal
    _fCy      : LREAL;                // 当拍有效周期 [s] / Effective cycle this scan
    _fPhStep  : LREAL;                // 相位单步上限 [deg] / Phase step ceiling
    _fScStep  : LREAL;                // 倍率单步上限 [%] / Scale step ceiling
    _bBusy    : BOOL := FALSE;        // 斜坡执行中内部量（R_TRIG 闸源） [-] / Busy internal
    _bClamped : BOOL;                 // 本拍应用沿发生钳位 [-] / Clamped at apply this scan
    _bRej     : BOOL;                 // 本拍应用沿被拒 [-] / Apply rejected this scan
    _bNonFin  : BOOL;                 // 请求非有限当拍量 [-] / Non-finite request this scan
    _bCfgBad  : BOOL;                 // 组态非法当拍量 [-] / Illegal configuration
    _bErrLatch: BOOL;                 // 组态故障锁存位（解除沿 = bReset 上升沿） / Latched config fault
    rtApply   : R_TRIG;               // 应用沿实例，段 0 无条件调用 / Apply edge instance
    rtReset   : R_TRIG;               // 复位沿实例，段 0 无条件调用 / Reset edge instance
END_VAR
VAR CONSTANT
    DL_CDT_CYDEF : LREAL := 0.01;     // 缺省扫描周期 [s] / Default scan cycle
    DL_CDT_TOL   : LREAL := 1.0E-9;   // 到达容差（禁浮点 = 判等） [deg|percent] / Arrival tolerance
    DL_CDT_ZERO  : LREAL := 0.0;      // 判零与安全侧基准 [deg|percent] / Zero base and safe value
    DL_CDT_UDMAX : UDINT := 4294967295;   // 拒次计数饱和点（防回绕） [次] / Reject counter ceiling
END_VAR

(* —— 段 0：非有限判 + 组态闸 + 周期派生 + 两沿无条件刷新 —— *)
_bNonFin := (fPhaseTrim <> fPhaseTrim) OR ((fPhaseTrim - fPhaseTrim) <> DL_CDT_ZERO)
         OR (fScaleTrim <> fScaleTrim) OR ((fScaleTrim - fScaleTrim) <> DL_CDT_ZERO);   // 请求非有限（R79 双判） / Non-finite request
_bCfgBad := (fPhTrimMaxDeg <= DL_CDT_ZERO) OR (fScTrimMaxPct <= DL_CDT_ZERO)
         OR (fPhRampDs <= DL_CDT_ZERO) OR (fScRampPs <= DL_CDT_ZERO)
         OR (fPhTrimMaxDeg <> fPhTrimMaxDeg) OR (fScTrimMaxPct <> fScTrimMaxPct);   // 组态域闸（上限/斜率域 + 上限非有限） / Configuration gate
IF fCycle > DL_CDT_ZERO THEN
    _fCy := fCycle;                   // 组态周期有效 / Configured cycle valid
ELSE
    _fCy := DL_CDT_CYDEF;             // 周期缺省兜底 / Default cycle fallback
END_IF
_fPhStep := fPhRampDs * _fCy;         // 相位单步 [deg] / Phase step
_fScStep := fScRampPs * _fCy;         // 倍率单步 [%] / Scale step
rtApply(CLK := bApply);               // 应用沿，每拍必调 / Apply edge, every scan
rtReset(CLK := bReset);               // 复位沿，每拍必调 / Reset edge, every scan

(* —— 段 1：复位沿与组态锁存 —— *)
IF rtReset.Q THEN
    _bErrLatch := FALSE;              // 清组态锁存（R188 声明：解除沿 = bReset 上升沿） / Clear cfg latch
    uRejCnt := 0;                     // 清拒次计数 / Clear reject counter
END_IF
IF _bCfgBad AND (NOT _bErrLatch) THEN
    _bErrLatch := TRUE;               // 锁存 / Latch
END_IF

(* —— 段 2：应用沿裁决（故障期拒绝；执行中拒绝叠加；请求钳位后锁存目标） —— *)
_bClamped := FALSE;                   // 钳位量预清 / Clamp preset
_bRej := FALSE;                       // 拒绝量预清 / Reject preset
IF rtApply.Q AND (NOT _bErrLatch) THEN
    IF _bBusy THEN
        _bRej := TRUE;                // 执行中拒绝叠加（规格，R191 声明：请求不生效，目标不变） / Busy reject, target unchanged
        IF uRejCnt < DL_CDT_UDMAX THEN
            uRejCnt := uRejCnt + 1;   // 拒次计数防回绕 / Count reject
        END_IF
    ELSIF _bNonFin THEN
        _bRej := TRUE;                // 非有限请求拒绝（不污染目标锁存） / Non-finite request rejected
        IF uRejCnt < DL_CDT_UDMAX THEN
            uRejCnt := uRejCnt + 1;   // 拒次计数 / Count reject
        END_IF
    ELSE
        _fPhTar := fPhaseTrim;        // 相位请求工作副本 / Phase working copy
        _fScTar := fScaleTrim;        // 倍率请求工作副本 / Scale working copy
        IF _fPhTar > fPhTrimMaxDeg THEN
            _fPhTar := fPhTrimMaxDeg;   // 相位超幅上钳（规格③） / Clamp phase high
            _bClamped := TRUE;          // 记钳位 / Mark clamp
        ELSIF _fPhTar < (-fPhTrimMaxDeg) THEN
            _fPhTar := -fPhTrimMaxDeg;  // 相位超幅下钳（对称 ±） / Clamp phase low
            _bClamped := TRUE;          // 记钳位 / Mark clamp
        END_IF
        IF _fScTar > fScTrimMaxPct THEN
            _fScTar := fScTrimMaxPct;   // 倍率超幅上钳 / Clamp scale high
            _bClamped := TRUE;          // 记钳位 / Mark clamp
        ELSIF _fScTar < (-fScTrimMaxPct) THEN
            _fScTar := -fScTrimMaxPct;  // 倍率超幅下钳 / Clamp scale low
            _bClamped := TRUE;          // 记钳位 / Mark clamp
        END_IF
        _bBusy := TRUE;               // 入斜坡执行态 / Enter ramp busy
    END_IF
END_IF

(* —— 段 3：双通道限步逼近（防凸轮表跳变；故障期冻结） —— *)
IF NOT _bErrLatch THEN
    IF _fPhTar > (_fPhAct + _fPhStep) THEN
        _fPhAct := _fPhAct + _fPhStep;   // 相位正向限步 / Phase ramp up
    ELSIF _fPhTar < (_fPhAct - _fPhStep) THEN
        _fPhAct := _fPhAct - _fPhStep;   // 相位负向限步 / Phase ramp down
    ELSE
        _fPhAct := _fPhTar;           // 相位步内到达 / Phase settle
    END_IF
    IF _fScTar > (_fScAct + _fScStep) THEN
        _fScAct := _fScAct + _fScStep;   // 倍率正向限步 / Scale ramp up
    ELSIF _fScTar < (_fScAct - _fScStep) THEN
        _fScAct := _fScAct - _fScStep;   // 倍率负向限步 / Scale ramp down
    ELSE
        _fScAct := _fScTar;           // 倍率步内到达 / Scale settle
    END_IF
    _bBusy := (ABS(_fPhAct - _fPhTar) >= DL_CDT_TOL)
           OR (ABS(_fScAct - _fScTar) >= DL_CDT_TOL);   // 双通道均达才撤销执行态（头注释④） / Busy until both settled
ELSE
    _bBusy := FALSE;                  // 故障期执行态强制撤销 / Fault forces not-busy
END_IF

(* —— 段 4：出口单点映射（名实双出口同源，R191） —— *)
fPhTrimAct := _fPhAct;                // 生效相位出口（故障期冻结保持） / Active phase outlet
fScTrimAct := _fScAct;                // 生效倍率出口 / Active scale outlet
bTrimActive := _bBusy;                // 执行中出口 / Busy outlet
IF _bErrLatch THEN
    bError := TRUE;                   // 故障标志（R45 配对） / Error flag
    eErrCode := E_DL_CdtErr.eCfgBad;  // 故障级码 / Fault code
ELSE
    bError := FALSE;                  // 无故障级条件 / No fault
    IF _bRej THEN
        eErrCode := E_DL_CdtErr.eBusyRej;   // 信息级：拒绝叠加 / Info: busy reject
    ELSIF _bClamped THEN
        eErrCode := E_DL_CdtErr.eClamped;   // 信息级：钳位口径 / Info: clamped
    ELSE
        eErrCode := E_DL_CdtErr.eOk;        // 正常 / Normal
    END_IF
END_IF

END_FUNCTION_BLOCK

(* ---- FB_DL_MultiAxisSyncErrGuard.st ---- *)
(*
    FB_DL_MultiAxisSyncErrGuard —— 多轴/龙门同步误差分级守护与首出诊断
    ------------------------------------------------------------------
    组件名    : FB_DL_MultiAxisSyncErrGuard
    分类      : DL_Motion / Synchronism Guard（多轴同步误差守护）
    一句话功能: 同时监控 4 个轴对的实时位置偏差，按「预警 → 降速 → 急停」三级响应，
                并在急停时锁存首出轴对编号与该对当时的误差值供诊断。
    复杂度    : C4
    版本      : v1.0.0
    开源溯源  : 无（clean-room 自研，未借鉴任何开源实现）
    平台      : 纯 IEC 61131-3（TON / R_TRIG / ABS / 标准库），目标编译器 RuSTy 1.0.8，
                兼容 CODESYS 3.5 / TwinCAT 3 / 汇川 InoProShop / Machine Expert；
                无 PROPERTY、无 VLA、无 FOR..DOWNTO、无厂商方言转换
    ------------------------------------------------------------------
    功能说明  : ① 每拍对 4 个轴对独立求同步误差 afErr[p] = ABS(afPosA[p] - afPosB[p])；
                ② 阈值三分：预警阈值 = fMaxSyncErrMm × fWarnRatio，
                   降速阈值 = fMaxSyncErrMm × fDerateRatio，急停阈值 = fMaxSyncErrMm；
                   组态闸强制 fWarnRatio < fDerateRatio < 1.0，故三带不交叠；
                ③ 建立窗口：使能有效后 tSettleMs 内不判误差（机构入位、伺服使能瞬态），
                   窗口未满只维持监控相，既不置预警也不置跳闸；
                ④ 降速相输出派生速度比例 fSpeedScalePct ∈ [50, 100]（单位 %），
                   比例随最大误差在「降速阈值 → 急停阈值」之间线性下降并饱和钳位；
                ⑤ 急停相 fSpeedScalePct = 0（安全侧：撤掉进给许可），并锁存首出轴对
                   编号与误差，供 HMI 直接定位是哪一对先越限；
                ⑥ 任一浮点输入为 NaN / ±Inf / 超幅值域 → 直接迁 eFault，bFaultOut := TRUE。
    量纲链    : afPosA [mm] − afPosB [mm] → afErr [mm]；
                fMaxSyncErrMm [mm] × fWarnRatio [-] → fThWarn [mm]（比例无因次，乘除不混加）；
                fMaxSyncErrMm [mm] × fDerateRatio [-] → fThDerate [mm]；
                (fWorstErr − fThDerate) [mm] ÷ (fMaxSyncErrMm − fThDerate) [mm] → fRto [-]
                （mm ÷ mm 无因次，符合线性归一）；
                fSpeedScalePct = 100 [%] − (100 − 50)[%] × fRto [-] → [%]；
                fFirstOutErr [mm] 原样输出不做任何换算。
                全程不存在「异量纲相加」：温度、时间、比例均不进入位置差的加法链。
    状态机    : eIdle(0) --使能且组态合法且输入有限--> eMonitor(10)
                eMonitor --nSev=1--> eWarn(20)
                eMonitor/eWarn --nSev=2--> eDerate(30)
                eMonitor/eWarn/eDerate --nSev=3（跳闸锁存）--> eTrip(40)
                eWarn --nSev=0--> eMonitor（逐级回落，无跨级跳跃）
                eDerate --nSev=1--> eWarn；--nSev=0--> eMonitor
                任意相 --非有限或组态非法--> eFault(90)
                eTrip / eFault 的唯一解除路径 = bReset 上升沿（见段 6 注释与自证行）
    失能语义  : bEnable = FALSE 时输出降级为安全值（eState := eIdle、fSpeedScalePct := 0、
                bWarn := FALSE），不冻结末值；bTrip / bFaultOut 锁存位不清 ——
                急停与故障必须人工复位，失能不能代替复位（安全侧口径，R191）。
    复位作用域: bReset 上升沿①清 _bTripLatch / _nFirstPair / _fFirstErr；
                ②清 _bFaultLatch 并迁相回 eIdle；③不清建立窗口锁存 _bSettled ——
                使能未断时保持「已建立」，避免复位后重新等窗口掩盖仍在恶化的偏差。
                复位沿与本拍跳闸同拍时：复位先执行、跳闸判断后执行，故本拍跳闸不被抹除
                （本拍合法事件优先，R275）。
    防御口径  : NaN 用自反 f<>f 判；±Inf 用 (f−f)<>(f−f) 双判；另设幅值域闸
                ABS(f) > 1.0E30 兜住超大有限值与 Inf 的观测域，三件套同拍生效（R4 + R151）。
                除零守卫：降速比例分母 (fMaxSyncErrMm − fThDerate) 先与 DL_SG_EPS 比较才做
                除法；组态闸另强制 fDerateRatio < 1.0，使分母结构性不小于
                fMaxSyncErrMm × (1 − fDerateRatio) > 0（双重保证，不靠单点）。
    规格偏离  : 派单输出引脚写作 iFirstOutPair（INT）。本库命名规范 1.2 规定有符号整数
                前缀为 n、i 专用于接口引用，故落为 nFirstOutPair，语义与取值范围
                （1..4，0 = 无首出）一字不减；另按 R190 归因唯一补充 bCfgErr / bDataErr
                两个诊断位，使「组态非法」与「数据非有限」两条故障成因各自可观测。
    码位说明  : 本件按零码位范式交付，不分配 16# 事件码；分级与故障一律经
                eState / bWarn / bTrip / bFaultOut / bCfgErr / bDataErr 组合观测。
    修订记录  : 2026-11-24 v1.0.0 首次入库（R87 批 · #1）
*)
TYPE E_DL_SyncState :
(
    eIdle    := 0,    // 空闲：未使能，速度比例锁 0，不判误差 | idle, disabled, speed scale forced to zero
    eMonitor := 10,   // 监控：使能且建立窗口已满，逐拍判误差，速度比例 100 | monitoring, window elapsed, scale 100
    eWarn    := 20,   // 预警：最大误差超预警阈值，限速不变，仅告警 | warning, threshold exceeded, speed unchanged
    eDerate  := 30,   // 降速：最大误差超降速阈值，速度比例按比例下降 | derate, speed scale ramped down
    eTrip    := 40,   // 急停：最大误差超上限，速度比例 0，首出轴对已锁存 | trip, scale zero, first-out latched
    eFault   := 90    // 故障：输入非有限或组态非法，锁存至复位沿 | fault latched until the reset edge
);
END_TYPE

FUNCTION_BLOCK FB_DL_MultiAxisSyncErrGuard
VAR_INPUT
    bEnable        : BOOL;                        // 使能电平，TRUE = 允许监控 | enable level, TRUE = monitoring allowed
    bReset         : BOOL;                        // 复位请求，上升沿生效 | reset request, rising-edge active
    afPosA         : ARRAY[1..4] OF REAL;         // 4 个轴对 A 侧实际位置 [mm] | actual position of the A side per pair [mm]
    afPosB         : ARRAY[1..4] OF REAL;         // 4 个轴对 B 侧实际位置 [mm] | actual position of the B side per pair [mm]
    fMaxSyncErrMm  : REAL := 1.0;                 // 同步误差上限（急停阈值）[mm] | sync error limit, trip threshold [mm]
    fWarnRatio     : REAL := 0.5;                 // 预警比例，乘上限得预警阈值 [-]，取值 (0,1) | warning ratio [dimensionless]
    fDerateRatio   : REAL := 0.8;                 // 降速比例，乘上限得降速阈值 [-]，取值 (warn,1) | derate ratio [dimensionless]
    tSettleMs      : TIME := T#200MS;             // 使能后的建立窗口，窗内不判 [ms] | settle window after enable [ms]
END_VAR
VAR_OUTPUT
    eState         : E_DL_SyncState;              // 主状态，供 HMI 与联锁使用 | main state for HMI and interlocks
    bWarn          : BOOL;                        // 预警汇总位，eWarn 或 eDerate 相为 TRUE | warning aggregate, TRUE in eWarn or eDerate
    bTrip          : BOOL;                        // 急停锁存位，复位沿前恒 TRUE | trip latch, stays TRUE until the reset edge
    fSpeedScalePct : REAL;                        // 派生速度比例指令 [%]，100 = 不限速，0 = 撤进给 | derived speed scale [%]
    nFirstOutPair  : INT;                         // 首出轴对编号 1..4，0 = 无首出 | first-out pair index 1..4, 0 = none
    fFirstOutErr   : REAL;                        // 首出轴对跳闸时的误差 [mm] | error of the first-out pair at trip [mm]
    bFaultOut      : BOOL;                        // 故障汇总位，含非有限与组态非法 | fault aggregate, covers non-finite and bad config
    bCfgErr        : BOOL;                        // 组态非法诊断位（归因唯一，R190）| bad-configuration flag, unique attribution
    bDataErr       : BOOL;                        // 数据非有限诊断位（归因唯一，R190）| non-finite data flag, unique attribution
END_VAR
VAR
    rtReset        : R_TRIG;                      // 复位上升沿实例，每拍无条件刷新 | reset rising-edge instance, refreshed every scan
    tonSettle      : TON;                         // 建立窗口计时实例，每拍无条件刷新 | settle window timer, refreshed every scan
    _eState        : E_DL_SyncState := E_DL_SyncState.eIdle; // 状态机内部当前态 | internal current state
    _bSettled      : BOOL := FALSE;               // 建立窗口已满锁存量 | settle-window elapsed latch
    _bResetLatch   : BOOL := FALSE;               // 复位沿锁存量，本拍末清除 | reset-edge latch, cleared at the end of the scan
    _bTripLatch    : BOOL := FALSE;               // 急停锁存位 | trip latch
    _bFaultLatch   : BOOL := FALSE;               // 故障锁存位 | fault latch
    _nFirstPair    : INT := 0;                    // 首出轴对编号锁存 1..4，0 = 无 | latched first-out pair index
    _fFirstErr     : REAL := 0.0;                 // 首出误差锁存 [mm] | latched first-out error [mm]
    afErr          : ARRAY[1..4] OF REAL;         // 各轴对同步误差绝对值 [mm] | absolute sync error per pair [mm]
    fThWarn        : REAL := 0.0;                 // 本拍预警阈值 [mm] | warning threshold this scan [mm]
    fThDerate      : REAL := 0.0;                 // 本拍降速阈值 [mm] | derate threshold this scan [mm]
    fWorstErr      : REAL := 0.0;                 // 本拍最大同步误差 [mm] | worst sync error this scan [mm]
    nWorstPair     : INT := 0;                    // 本拍最大误差所属轴对 1..4 | pair holding the worst error this scan
    nTripPair      : INT := 0;                    // 本拍首个越急停阈值的轴对 1..4 | lowest-index pair beyond the trip threshold
    nSev           : INT := 0;                    // 本拍严重度 0 正常 1 预警 2 降速 3 急停 | severity level this scan
    nIdx           : INT := 1;                    // 轴对遍历下标 | pair loop index
    _bBadIn        : BOOL := FALSE;               // 本拍输入非有限标志 | non-finite input flag this scan
    _bCfgBad       : BOOL := FALSE;               // 本拍组态非法标志 | bad configuration flag this scan
    fDen           : REAL := 0.0;                 // 降速比例分母（阈值带宽）[mm] | derate scaling denominator [mm]
    fRto           : REAL := 0.0;                 // 降速带内归一比例 [0..1] | normalised ratio inside the derate band
END_VAR
VAR CONSTANT
    DL_SG_PAIR_MAX   : INT := 4;                  // 轴对总数硬界，与数组上界一致 [-] | hard pair count matching the array bound
    DL_SG_EPS        : REAL := 1.0E-6;            // 浮点判零容差 [mm] | float zero tolerance [mm]
    DL_SG_MAG_MAX    : REAL := 1.0E30;            // 有限幅值域闸上限 [mm] | finite magnitude domain bound [mm]
    DL_SG_SCALE_MIN  : REAL := 50.0;              // 降速相最低速度比例 [%] | minimum derated speed scale [%]
    DL_SG_SCALE_FULL : REAL := 100.0;             // 满速比例 [%] | full speed scale [%]
END_VAR

METHOD Clamp01 : REAL
(*
    归一比例钳位：把降速带内比例钳到 [0,1]，越界一律饱和。纯函数，无跨拍状态。
    Clamp-normalised ratio: saturate the in-band ratio to [0,1]. Pure function, no cross-scan state.
*)
VAR_INPUT
    fIn : REAL;                                   // 待钳位比例 [-] | ratio to be clamped [-]
END_VAR
Clamp01 := fIn;                                   // 直通赋值，下方按两侧硬界饱和 | straight-through, saturated on both bounds below
IF Clamp01 < 0.0 THEN
    Clamp01 := 0.0;                               // 低于下限钳 0，防负比例抬高速度 | clamp low bound to zero
END_IF
IF Clamp01 > 1.0 THEN
    Clamp01 := 1.0;                               // 高于上限钳 1，防比例超上限 | clamp high bound to one
END_IF
END_METHOD

// 段 1｜定时器与沿实例无条件周期刷新（R7：严禁放入 IF / CASE 分支内部）
// segment 1, timers and edge instances refreshed unconditionally, never inside an IF or CASE branch
rtReset(CLK := bReset);
tonSettle(IN := bEnable AND (NOT _bSettled), PT := tSettleMs);
IF rtReset.Q THEN
    _bResetLatch := TRUE;                         // 复位沿先存锁存量，由段 6 统一消费 | store the reset edge, consumed in segment 6
END_IF
IF tonSettle.Q THEN
    _bSettled := TRUE;                            // 窗口到时置锁存量，本拍即可判 | window elapsed, judging allowed from this scan
END_IF
IF NOT bEnable THEN
    _bSettled := FALSE;                           // 失能即重新武装窗口，下次使能重新计时 | disarm the window so the next enable re-times
END_IF

// 段 2｜输出安全侧预置（每拍先落安全值，CASE 内只做升级赋值）
// segment 2, preset outputs to their safe values; the CASE below only upgrades them
fSpeedScalePct := 0.0;                            // 预置速度比例 0 [%]，进给许可默认撤销 | preset zero speed scale, feed permission withdrawn
bWarn := FALSE;                                   // 预置无预警 | preset no warning
_bBadIn := FALSE;                                 // 预置输入有限 | preset finite input
_bCfgBad := FALSE;                                // 预置组态合法 | preset legal configuration
nSev := 0;                                        // 预置严重度正常 | preset normal severity

// 段 3｜非有限闸：NaN 自反 + Inf 自减 + 幅值域，逐个浮点入参枚举（R4 / R151 / R272）
// segment 3, non-finite gate: NaN self-reflexive, Inf by self-subtraction, plus a magnitude bound, one entry per REAL input
FOR nIdx := 1 TO DL_SG_PAIR_MAX DO
    IF (afPosA[nIdx] <> afPosA[nIdx]) OR ((afPosA[nIdx] - afPosA[nIdx]) <> (afPosA[nIdx] - afPosA[nIdx])) THEN
        _bBadIn := TRUE;                          // A 侧 NaN 或 ±Inf | NaN or infinity on the A side
    END_IF
    IF ABS(afPosA[nIdx]) > DL_SG_MAG_MAX THEN
        _bBadIn := TRUE;                          // A 侧超幅值域 | A side beyond the magnitude domain
    END_IF
    IF (afPosB[nIdx] <> afPosB[nIdx]) OR ((afPosB[nIdx] - afPosB[nIdx]) <> (afPosB[nIdx] - afPosB[nIdx])) THEN
        _bBadIn := TRUE;                          // B 侧 NaN 或 ±Inf | NaN or infinity on the B side
    END_IF
    IF ABS(afPosB[nIdx]) > DL_SG_MAG_MAX THEN
        _bBadIn := TRUE;                          // B 侧超幅值域 | B side beyond the magnitude domain
    END_IF
END_FOR
IF (fMaxSyncErrMm <> fMaxSyncErrMm) OR ((fMaxSyncErrMm - fMaxSyncErrMm) <> (fMaxSyncErrMm - fMaxSyncErrMm)) THEN
    _bBadIn := TRUE;                              // 误差上限 NaN 或 ±Inf | limit NaN or infinity
END_IF
IF (fWarnRatio <> fWarnRatio) OR ((fWarnRatio - fWarnRatio) <> (fWarnRatio - fWarnRatio)) THEN
    _bBadIn := TRUE;                              // 预警比例 NaN 或 ±Inf | warning ratio NaN or infinity
END_IF
IF (fDerateRatio <> fDerateRatio) OR ((fDerateRatio - fDerateRatio) <> (fDerateRatio - fDerateRatio)) THEN
    _bBadIn := TRUE;                              // 降速比例 NaN 或 ±Inf | derate ratio NaN or infinity
END_IF

// 段 4｜组态闸：上限须为正、比例须严格递增且小于 1（保证三带不交叠、降速分母为正）
// segment 4, configuration gate: positive limit, strictly increasing ratios below one, keeping three disjoint bands and a positive denominator
IF (fMaxSyncErrMm <= DL_SG_EPS) OR (fWarnRatio <= DL_SG_EPS) OR (fWarnRatio >= fDerateRatio) OR (fDerateRatio >= 1.0) THEN
    _bCfgBad := TRUE;                             // 组态非法：阈值带错序或非正 | illegal configuration, band order or sign
END_IF

// 段 5｜阈值、误差与严重度裁决（每拍全量重算，无跨拍状态驻留）
// segment 5, thresholds, errors and severity decision, fully recomputed every scan with no cross-scan state
fThWarn := fMaxSyncErrMm * fWarnRatio;            // 预警阈值 [mm] = [mm] × [-] | warning threshold [mm]
fThDerate := fMaxSyncErrMm * fDerateRatio;        // 降速阈值 [mm] = [mm] × [-] | derate threshold [mm]
fWorstErr := 0.0;                                 // 清本拍最大误差 [mm] | clear the worst error
nWorstPair := 0;                                  // 清本拍最坏轴对编号 | clear the worst pair index
nTripPair := 0;                                   // 清本拍首个越限轴对编号 | clear the lowest-index tripping pair
FOR nIdx := 1 TO DL_SG_PAIR_MAX DO
    afErr[nIdx] := ABS(afPosA[nIdx] - afPosB[nIdx]); // 轴对同步误差 [mm] = [mm] − [mm] | per-pair sync error [mm]
    IF afErr[nIdx] > fWorstErr THEN
        fWorstErr := afErr[nIdx];                 // 记录本拍最大误差 [mm] | record the worst error [mm]
        nWorstPair := nIdx;                       // 记录最大误差所属轴对 | record the pair holding it
    END_IF
    IF (afErr[nIdx] > fMaxSyncErrMm) AND (nTripPair = 0) THEN
        nTripPair := nIdx;                        // 升序遍历只记首个越限对，首出不随最坏值漂移 | first tripping pair only, ascending scan
    END_IF
END_FOR
IF fWorstErr > fMaxSyncErrMm THEN
    nSev := 3;                                    // 超急停上限 | beyond the trip limit
ELSIF fWorstErr > fThDerate THEN
    nSev := 2;                                    // 超降速阈值 | beyond the derate threshold
ELSIF fWorstErr > fThWarn THEN
    nSev := 1;                                    // 超预警阈值 | beyond the warning threshold
ELSE
    nSev := 0;                                    // 三带之内正常运行 | inside all bands, normal operation
END_IF

// 段 6｜复位沿处理（唯一解除路径）：先复位后判跳闸，保证本拍新跳闸不被抹除（R275）
// segment 6, reset edge handling, the only release path; reset runs before the trip decision so a same-scan trip survives
IF _bResetLatch THEN
    _bTripLatch := FALSE;                         // 清急停锁存 | clear the trip latch
    _nFirstPair := 0;                             // 清首出轴对编号 | clear the first-out pair index
    _fFirstErr := 0.0;                            // 清首出误差 [mm] | clear the first-out error [mm]
    _bFaultLatch := FALSE;                        // 清故障锁存 | clear the fault latch
    _eState := E_DL_SyncState.eIdle;              // 迁回空闲相，下一拍按使能重新建窗 | return to idle, re-arm on the next scan
END_IF

// 段 7｜故障锁存：非有限与组态非法各自独立置位（R190 归因唯一），锁存与迁相同段完成
// segment 7, fault latches; non-finite data and bad configuration keep separate members and separate set points
IF _bBadIn AND (NOT _bFaultLatch) THEN
    _bFaultLatch := TRUE;                         // 锁存数据非有限 | latch the non-finite data fault
    _eState := E_DL_SyncState.eFault;             // 与锁存同拍迁相（R258）| migrate in the same scan as the latch
END_IF
IF _bCfgBad AND (NOT _bFaultLatch) THEN
    _bFaultLatch := TRUE;                         // 锁存组态非法 | latch the bad configuration fault
    _eState := E_DL_SyncState.eFault;             // 与锁存同拍迁相（R258）| migrate in the same scan as the latch
END_IF

// 段 8｜跳闸判据与首出锁存：与状态无关的纯判据，故放在 CASE 之前统一裁决
// segment 8, trip criterion and first-out latch; a state-independent criterion, so it is decided before the CASE
IF bEnable AND _bSettled AND (NOT _bTripLatch) AND (NOT _bFaultLatch) AND (nSev >= 3) THEN
    _bTripLatch := TRUE;                          // 置急停锁存 | raise the trip latch
    IF nTripPair > 0 THEN
        _nFirstPair := nTripPair;                 // 首出 = 首个越限轴对 | first out is the lowest-index tripping pair
    ELSE
        _nFirstPair := nWorstPair;                // 兜底取最坏轴对（结构上 nSev>=3 必有越限对）| fall back to the worst pair
    END_IF
    _fFirstErr := fWorstErr;                      // 记录当时误差 [mm] | record the error at trip [mm]
END_IF

// 段 9｜主状态机：ENUM + CASE + ELSE 兜底（R6），逐级升降，无跨级跳跃
// segment 9, main state machine with ENUM + CASE + ELSE fallback, stepwise up and down, no band skipping
CASE _eState OF
E_DL_SyncState.eIdle:
    fSpeedScalePct := 0.0;                        // 空闲相速度比例 0 [%] | idle phase keeps the scale at zero
    // 拍 N 进入：复位沿或使能撤除；本拍行为：拒绝任何分级输出，只保留锁存位；
    // 拍 N+1 转出：使能有效且组态合法且输入有限 → 监控相
    // entered on the reset edge or on disable; refuses every graded output and keeps the latches only;
    // exits to eMonitor once enabled with legal configuration and finite inputs
    IF bEnable AND (NOT _bCfgBad) AND (NOT _bBadIn) AND (NOT _bFaultLatch) THEN
        _eState := E_DL_SyncState.eMonitor;
    END_IF

E_DL_SyncState.eMonitor:
    fSpeedScalePct := DL_SG_SCALE_FULL;           // 监控相满速 100 [%] | monitoring phase runs at full scale [%]
    IF NOT bEnable THEN
        _eState := E_DL_SyncState.eIdle;           // 失能回空闲 | return to idle when disabled
    ELSIF _bTripLatch THEN
        _eState := E_DL_SyncState.eTrip;           // 本拍跳闸优先迁移 | migrate to trip when the latch is raised
    ELSIF _bSettled AND (nSev = 2) THEN
        _eState := E_DL_SyncState.eDerate;         // 升到降速相 | step up to derate
    ELSIF _bSettled AND (nSev = 1) THEN
        _eState := E_DL_SyncState.eWarn;           // 升到预警相 | step up to warning
    END_IF
    // 窗口未满时不迁移也不降级：偏差在建立窗口内无意义 | inside the settle window no migration is taken, deviation is meaningless there

E_DL_SyncState.eWarn:
    fSpeedScalePct := DL_SG_SCALE_FULL;           // 预警相不限速 100 [%] | warning phase keeps full scale [%]
    IF NOT bEnable THEN
        _eState := E_DL_SyncState.eIdle;           // 失能回空闲 | return to idle when disabled
    ELSIF _bTripLatch THEN
        _eState := E_DL_SyncState.eTrip;           // 急停优先 | trip takes priority
    ELSIF (NOT _bSettled) THEN
        _eState := E_DL_SyncState.eMonitor;        // 窗口被重新武装（使能曾断）→ 回监控等窗口 | window re-armed, wait in monitoring
    ELSIF nSev = 2 THEN
        _eState := E_DL_SyncState.eDerate;         // 恶化升相 | worsen to derate
    ELSIF nSev = 0 THEN
        _eState := E_DL_SyncState.eMonitor;        // 回落到正常带 → 降相 | back inside the bands, step down
    END_IF

E_DL_SyncState.eDerate:
    // 降速比例：误差在「降速阈值 → 急停阈值」之间线性下降到 DL_SG_SCALE_MIN [%]
    // derate scale: linear descent from the derate threshold to the trip limit, saturating at the minimum scale
    fDen := fMaxSyncErrMm - fThDerate;            // 降速带宽 [mm] = [mm] − [mm] | derate band width [mm]
    IF fDen > DL_SG_EPS THEN
        fRto := Clamp01((fWorstErr - fThDerate) / fDen); // 带内归一比例 [-] = [mm] ÷ [mm]，先判零再除 | guarded division
    ELSE
        fRto := 1.0;                              // 分母为零宽（组态闸已禁）→ 保守取满比例 | degenerate width, take the saturated ratio
    END_IF
    fSpeedScalePct := DL_SG_SCALE_FULL - (DL_SG_SCALE_FULL - DL_SG_SCALE_MIN) * fRto; // [%] − [%] × [-] | derated scale [%]
    IF NOT bEnable THEN
        _eState := E_DL_SyncState.eIdle;           // 失能回空闲 | return to idle when disabled
    ELSIF _bTripLatch THEN
        _eState := E_DL_SyncState.eTrip;           // 急停优先 | trip takes priority
    ELSIF (NOT _bSettled) THEN
        _eState := E_DL_SyncState.eMonitor;        // 窗口重新武装 → 回监控 | window re-armed, wait in monitoring
    ELSIF nSev >= 3 THEN
        _eState := E_DL_SyncState.eTrip;           // 越急停上限（锁存同拍已置）| beyond the trip limit, latch already raised
    ELSIF nSev = 0 THEN
        _eState := E_DL_SyncState.eMonitor;        // 直接回到正常带 | straight back to the normal band
    ELSIF nSev = 1 THEN
        _eState := E_DL_SyncState.eWarn;           // 缓解到预警带 | relieved into the warning band
    END_IF

E_DL_SyncState.eTrip:
    fSpeedScalePct := 0.0;                        // 急停相速度比例 0 [%]，撤进给许可 | trip phase withdraws the feed permission
    // 驻留语义：本相只能由段 6 复位沿迁出（唯一解除路径），本相不再判误差
    // dwell semantics: this phase is left only through the reset edge handled in segment 6, no error judging here

E_DL_SyncState.eFault:
    fSpeedScalePct := 0.0;                        // 故障相速度比例 0 [%] | fault phase withdraws the feed permission
    // 驻留语义：本相只能由段 6 复位沿迁出；故障码由 _bBadIn / _bCfgBad 分别观测（R190）
    // dwell semantics: left only through the reset edge in segment 6; causes observed via _bBadIn and _bCfgBad separately

ELSE
    // 非法枚举值（越界或未定义成员）：不猜、不驻留，直接置故障并回故障相
    // illegal enumerator: no guessing, latch a fault and return to the fault phase
    fSpeedScalePct := 0.0;
    _bFaultLatch := TRUE;
    _eState := E_DL_SyncState.eFault;
END_CASE;

// 段 10｜出口单点映射（锁存位在本段回放，CASE 后不再无条件清零任何 CASE 内写过的量，R187）
// segment 10, single-point output mapping; latches are replayed here and nothing written inside the CASE is cleared afterwards
eState := _eState;                                // 状态映射 | state mapping
bWarn := (_eState = E_DL_SyncState.eWarn) OR (_eState = E_DL_SyncState.eDerate); // 预警汇总，由状态派生 | warning derived from the state
bTrip := _bTripLatch;                             // 急停锁存回放 | replay the trip latch
bFaultOut := _bFaultLatch;                        // 故障锁存回放 | replay the fault latch
bCfgErr := _bCfgBad;                              // 组态非法诊断位 | bad-configuration diagnostic
bDataErr := _bBadIn;                              // 数据非有限诊断位 | non-finite data diagnostic
nFirstOutPair := _nFirstPair;                     // 首出轴对编号回放 | replay the first-out pair index
fFirstOutErr := _fFirstErr;                       // 首出误差回放 [mm] | replay the first-out error [mm]

// 段 11｜本拍消费量收尾（仅清沿锁存，不触碰任何锁存位与 CASE 内写入量）
// segment 11, end-of-scan cleanup; only the edge latch is cleared, no latch and no CASE-written identifier is touched
_bResetLatch := FALSE;
END_FUNCTION_BLOCK
